			IF Munsch.bSetAirTemp
			THEN
				nWatchdog := 0;
				bDone:= FALSE;                               		(* Program done *)
				bBusy := TRUE;                                  	(* Program busy *)
	
				Munsch.bLockedInterface := TRUE;
				Munsch.bSendExe := FALSE;
	
				IF nAirTemp >= nMinAirTemp
				     AND nAirTemp <= nMaxAirTemp
				THEN
					etMunschExtruder := ET_MunschExtruder_eSetCMD;              (* Next step *)
				ELSE
					udnErrorNo := 1;
	
					etMunschExtruder := ET_MunschExtruder_eError;              (* Next step *)
				END_IF

			ELSE
				etMunschExtruder := ET_MunschExtruder_eError;             (* Next step *)
			END_IF

			Munsch.bSetAirTemp := FALSE;

		ELSIF nWatchdog > 1000
		THEN
			Munsch.bSetAirTemp := FALSE;

			etMunschExtruder := ET_MunschExtruder_eError;             (* Next step *)
		END_IF

	ET_MunschExtruder_eSetCMD:
		Munsch.stMunschCmd.etCommand := ET_MUNSCH_CMD_SETAIRTEMP;
		Munsch.stMunschCmd.nAirTemp := nAirTemp;

		etMunschExtruder := ET_MunschExtruder_eExecuteCMD;              (* Next step *)

	ET_MunschExtruder_eExecuteCMD:
		nWatchdog := nWatchdog + 1;

		Munsch.bSendExe := TRUE;

		IF Munsch.bStringReceived
		THEN
			IF Munsch.stMunschRes.etResponse = ET_MUNSCH_RES_SETAIRTEMP
			     AND Munsch.stMunschCmd.nAirTemp = Munsch.stMunschRes.nAirRefTemp
			THEN
				Munsch.bSendExe := FALSE;

				nWatchdog := 0;

				etMunschExtruder := ET_MunschExtruder_eSetREQ;              (* Next step *)

			END_IF

		ELSIF Munsch.bInterfaceError
			    OR nWatchdog > 1000
		THEN
			Munsch.bSendExe := FALSE;

			udnErrorNo := 2;                     (* Error number *)
			etMunschExtruder := ET_MunschExtruder_eError;              (* Next step *)

		END_IF

	ET_MunschExtruder_eSetREQ:
		Munsch.stMunschCmd.etCommand := ET_MUNSCH_CMD_REQAIRREFTEMP;

		etMunschExtruder := ET_MunschExtruder_eExecuteREQ;              (* Next step *)

	ET_MunschExtruder_eExecuteREQ:
		nWatchdog := nWatchdog + 1;

		Munsch.bSendExe := TRUE;

		IF Munsch.bStringReceived
		THEN
			IF Munsch.stMunschRes.etResponse = ET_MUNSCH_RES_REQAIRREFTEMP
			THEN
				Munsch.nAirRefTemp := Munsch.stMunschRes.nAirRefTemp;

				Munsch.bSendExe := FALSE;

				nWatchdog := 0;
				etMunschExtruder := ET_MunschExtruder_eDone;              (* Next step *)
			END_IF

		ELSIF Munsch.bInterfaceError
			    OR nWatchdog > 1000
		THEN
			Munsch.bSendExe := FALSE;

			udnErrorNo := 3;                     (* Error number *)
			etMunschExtruder := ET_MunschExtruder_eError;              (* Next step *)

		END_IF

	ET_MunschExtruder_eError:
		bBusy := FALSE;						(* Command busy *)
		bError := TRUE;						(* Command error  *)

		etMunschExtruder := ET_MunschExtruder_eNoExecute;

	ET_MunschExtruder_eDone:
		bDone := TRUE;						(* Command done *)
		bBusy := FALSE;						(* Command busy *)

		etMunschExtruder := ET_MunschExtruder_eNoExecute;

	ET_MunschExtruder_eNoExecute:
		IF NOT bExecute
		THEN
			(* Reset outputs *)
			bDone := FALSE;						(* Command done *)
			bBusy := FALSE;						(* Command busy *)
			bError := FALSE;						(* Command error  *)

			nWatchdog := 0;
			Munsch.bLockedInterface := FALSE;

			Munsch.stMunschCmd.etCommand := ET_MUNSCH_CMD_NOCMD;
			Munsch.stMunschRes.etResponse := ET_MUNSCH_RES_NOCMD;

			etMunschExtruder := ET_MunschExtruder_eWaitExecute;
		END_IF
END_CASE;

bAirTempAlarm := Munsch.nAirActTemp > Munsch.nAirRefTemp + nAirTempTolerance
				OR Munsch.nAirActTemp > Munsch.nAirRefTemp - nAirTempTolerance;

END_FUNCTION_BLOCK

// ---- POUs/Tc2 Objects/ExternalHardware/Munsch/FB_MunschExtruder_Extruding.TcPOU
FUNCTION_BLOCK FB_MunschExtruder_Extruding
(*

The function block used to control extruding Munsch extruder

Constructor: 		Patryk Panylo
Company:		E. Riexinger GmbH
Date:			13.10.2015
Version:			1.00

Date:			Revision:		Who:				Comment
dd.mm.yyyy		x.xx			Initials			comment

*)
VAR_INPUT
	(* Input variables / Eingang Variablen *)
	bEnable						:BOOL;						(* Enable FB signal *)
	bStart						:BOOL;						(* Start heating *)
	bStop						:BOOL;						(* Start heating *)
	nExtrudingSpeed				:INT;						(* Extruding speed [%] *)
	rExtrudingSpeedOffset			:REAL;						(* Extruding speed [%] *)
	lrExtrudingSpeedMinV			:LREAL;						(* Extruding speed min [V] 16#0000 = 0 [V] *)
	lrExtrudingSpeedMaxV 		:LREAL;						(* Extruding speed max [V] 16#7FFF = 10 [V], 16#3FFF = 5[V] *)
	lrExtrudingSpeedMin			:LREAL;						(* Extruding speed min [%] *)
	lrExtrudingSpeedMax			:LREAL;						(* Extruding speed max [%] *)
END_VAR
VAR_OUTPUT
	(* Output variables / Ausgang Variablen *)
	bDone						:BOOL;						(* Program done *)
	bBusy						:BOOL;						(* Program busy *)
	bError						:BOOL;						(* Error *)
	udnErrorNo					:UDINT;
END_VAR
VAR_IN_OUT
	(* Input Output variables / Ausgang Variablen *)
	Munsch						:ST_MUNSCH_REF;
END_VAR
VAR
	(* Enummerations *)
	etMunschExtruder				:ET_MunschExtruder;

	(* Variables *)
	nWatchdog					:INT;

	nExtrudingSpeedLimitMax		:INT := 16383;					(* The extruding speed limit (absolute value). Value range in V: 0 ...10, 16#3FFF = 5[V]*)

	(* References *)

	(* Interfaces *)

	(* Instances *)
	fbExtrudingSpeed				:FB_ScalingOffset;
	rtStart						:R_TRIG;
	rtStop						:R_TRIG;

	rtStartEx						:R_TRIG;
	rtStopEx						:R_TRIG;
	bStartEx						:BOOL;
	bStopEx						:BOOL;
END_VAR

IF NOT bEnable
THEN
	bDone := FALSE;					(* Program done *)
	bBusy := FALSE;                                  	(* Program not busy *)
	bError := FALSE;                                 	(* Program not error *)
	udnErrorNo := 0;                                 		(* Error number *)

	Munsch.bExtruding := FALSE;

	RETURN;
END_IF;

(* Scale extruding speed *)
fbExtrudingSpeed(
	bEnable := TRUE,
	lrInput := INT_TO_LREAL(nExtrudingSpeed),
	lrXLowLimit := lrExtrudingSpeedMin,
	lrXUpperLimit := lrExtrudingSpeedMax,
	lrYLowLimit := lrExtrudingSpeedMinV,
	lrYUpperLimit := MIN(lrExtrudingSpeedMaxV, nExtrudingSpeedLimitMax),
	usiPrecision := 2,
	lrOffset := rExtrudingSpeedOffset
);

IF NOT Munsch.bHeat
     OR NOT Munsch.bHeated
     OR NOT Munsch.bExtruding
THEN
	Munsch.nExtrudingSpeed := 0;
	(*bStartEx := FALSE;
	bStopEx := FALSE;*)
ELSE
	(*Munsch.nExtrudingSpeed := LREAL_TO_INT(fbExtrudingSpeed.lrOutputPV);*);
END_IF

(* Wait for triger *)
rtStart(
	CLK := bStart
);

rtStop(
	CLK := bStop
);

(* Wait for triger *)
rtStartEx(
	CLK := Munsch.stMunschCmd.etCommand = ET_MUNSCH_CMD_STARTEXTRUDER
		    AND Munsch.stMunschRes.etResponse = ET_MUNSCH_RES_STARTEXTRUDER
		    AND bBusy
);

rtStopEx(
	CLK := Munsch.stMunschCmd.etCommand = ET_MUNSCH_CMD_STOPEXTRUDER
	  	    AND Munsch.stMunschRes.etResponse = ET_MUNSCH_RES_STOPEXTRUDER
		    AND bBusy
);

IF rtStopEx.Q
THEN
	bStartEx := FALSE;
	bStopEx := TRUE;

ELSIF rtStartEx.Q
THEN
	bStartEx := TRUE;
	bStopEx := FALSE;

END_IF

IF bStopEx
THEN
	Munsch.nExtrudingSpeed := 0;
ELSIF bStartEx
THEN
	Munsch.nExtrudingSpeed := LREAL_TO_INT(fbExtrudingSpeed.lrOutputPV);
END_IF

IF rtStop.Q
THEN
	Munsch.bSetAirTemp := FALSE;
	Munsch.bSetMaterialTemp := FALSE;
	Munsch.bStartHeat := FALSE;
	Munsch.bStopHeat  := FALSE;
	Munsch.bStartExtruding := FALSE;
	Munsch.bStopExtruding  := TRUE;
	Munsch.bReadStatus := FALSE;

	Munsch.nExtrudingSpeed := 0;
END_IF

(* Send command *)
CASE etMunschExtruder OF

	ET_MunschExtruder_eWaitExecute:
		IF rtStop.Q
		    OR Munsch.bStopExtruding
		    OR (nExtrudingSpeed = 0
			   AND Munsch.bExtruding)
		THEN
			nWatchdog := 0;

			Munsch.bSetAirTemp := FALSE;
			Munsch.bSetMaterialTemp := FALSE;
			Munsch.bStartHeat := FALSE;
			Munsch.bStopHeat  := FALSE;
			Munsch.bStartExtruding := FALSE;
			Munsch.bStopExtruding  := TRUE;
			Munsch.bReadStatus := FALSE;

			Munsch.nExtrudingSpeed := 0;

			etMunschExtruder := ET_MunschExtruder_eChkInterface;              (* Next step *)

		ELSIF rtStart.Q
		    	    AND Munsch.bHeat
		             AND Munsch.bHeated
		THEN
			nWatchdog := 0;

			Munsch.bSetAirTemp := FALSE;
			Munsch.bSetMaterialTemp := FALSE;
			Munsch.bStartHeat := FALSE;
			Munsch.bStopHeat  := FALSE;
			Munsch.bStartExtruding := TRUE;
			Munsch.bStopExtruding  := FALSE;
			Munsch.bReadStatus := FALSE;

			etMunschExtruder := ET_MunschExtruder_eChkInterface;              (* Next step *)

		END_IF

	ET_MunschExtruder_eChkInterface:
		nWatchdog := nWatchdog + 1;

		IF NOT Munsch.bLockedInterface
		THEN
			bBusy := FALSE;                                     	(* Program not busy *)
			bError := FALSE;                         		(* Program not error *)
			udnErrorNo := 0;                         		(* Error number *)

			IF Munsch.bStopExtruding
			THEN
				nWatchdog := 0;
				bDone:= FALSE;                               		(* Program done *)
				bBusy := TRUE;                                  	(* Program busy *)
	
				Munsch.nExtrudingSpeed := 0;
	
				Munsch.bLockedInterface := TRUE;
				Munsch.bSendExe := FALSE;
				Munsch.stMunschCmd.etCommand := ET_MUNSCH_CMD_STOPEXTRUDER;
	
				etMunschExtruder := ET_MunschExtruder_eSetCMD;              (* Next step *)
	
			ELSIF Munsch.bStartExtruding
			THEN
				nWatchdog := 0;
				bDone:= FALSE;                               		(* Program done *)
				bBusy := TRUE;                                  	(* Program busy *)
	
				Munsch.nExtrudingSpeed := LREAL_TO_INT(fbExtrudingSpeed.lrOutputPV);
	
				Munsch.bLockedInterface := TRUE;
				Munsch.bSendExe := FALSE;
				Munsch.stMunschCmd.etCommand := ET_MUNSCH_CMD_STARTEXTRUDER;
	
				etMunschExtruder := ET_MunschExtruder_eSetCMD;              (* Next step *)

			ELSE
				etMunschExtruder := ET_MunschExtruder_eError;             (* Next step *)
			END_IF

			Munsch.bStartExtruding := FALSE;
			Munsch.bStopExtruding  := FALSE;

		ELSIF nWatchdog > 1000
		THEN
			Munsch.bStartExtruding := FALSE;
			Munsch.bStopExtruding  := FALSE;

			etMunschExtruder := ET_MunschExtruder_eError;             (* Next step *)
		END_IF

	ET_MunschExtruder_eSetCMD:
		etMunschExtruder := ET_MunschExtruder_eExecuteCMD;              (* Next step *)

	ET_MunschExtruder_eExecuteCMD:
		nWatchdog := nWatchdog + 1;

		Munsch.bSendExe := TRUE;

		IF Munsch.bStringReceived
		THEN
			IF (Munsch.stMunschCmd.etCommand = ET_MUNSCH_CMD_STARTEXTRUDER
			      AND Munsch.stMunschRes.etResponse = ET_MUNSCH_RES_STARTEXTRUDER)
			     OR
			     (Munsch.stMunschCmd.etCommand = ET_MUNSCH_CMD_STOPEXTRUDER
			      AND Munsch.stMunschRes.etResponse = ET_MUNSCH_RES_STOPEXTRUDER)
			THEN
				Munsch.bSendExe := FALSE;

				nWatchdog := 0;
				etMunschExtruder := ET_MunschExtruder_eSetREQ;              (* Next step *)

			END_IF

		ELSIF Munsch.bInterfaceError
			    OR nWatchdog > 1000
		THEN
			Munsch.bSendExe := FALSE;

			udnErrorNo := 1;                     (* Error number *)

			etMunschExtruder := ET_MunschExtruder_eError;              (* Next step *)
		END_IF

	ET_MunschExtruder_eSetREQ:
		Munsch.stMunschCmd.etCommand := ET_MUNSCH_CMD_REQEXTRUDERSTATUS;

		etMunschExtruder := ET_MunschExtruder_eExecuteREQ;              (* Next step *)

	ET_MunschExtruder_eExecuteREQ:
		nWatchdog := nWatchdog + 1;

		Munsch.bSendExe := TRUE;

		IF Munsch.bStringReceived
		THEN
			IF Munsch.stMunschRes.etResponse = ET_MUNSCH_RES_ACKEXTRUDERSTATUSON
			THEN
				Munsch.bExtruding := TRUE;
				Munsch.bSendExe := FALSE;

				nWatchdog := 0;
				etMunschExtruder := ET_MunschExtruder_eDone;              (* Next step *)
			
			ELSIF Munsch.stMunschRes.etResponse = ET_MUNSCH_RES_ACKEXTRUDERSTATUSOFF
			THEN
				Munsch.bExtruding := FALSE;
				Munsch.bSendExe := FALSE;

				nWatchdog := 0;
				etMunschExtruder := ET_MunschExtruder_eDone;              (* Next step *)

			END_IF

		ELSIF Munsch.bInterfaceError
			    OR nWatchdog > 1000
		THEN
			Munsch.bSendExe := FALSE;

			udnErrorNo := 2;                     (* Error number *)

			etMunschExtruder := ET_MunschExtruder_eError;              (* Next step *)
		END_IF

	ET_MunschExtruder_eError:
		bBusy := FALSE;						(* Command busy *)
		bError := TRUE;						(* Command error  *)

		etMunschExtruder := ET_MunschExtruder_eNoExecute;

	ET_MunschExtruder_eDone:
		bDone := TRUE;						(* Command done *)
		bBusy := FALSE;						(* Command busy *)

		etMunschExtruder := ET_MunschExtruder_eNoExecute;

	ET_MunschExtruder_eNoExecute:
		IF NOT bStart
		     AND NOT bStop
		THEN
			(* Reset outputs *)
			bDone := FALSE;						(* Command done *)
			bBusy := FALSE;						(* Command busy *)
			bError := FALSE;						(* Command error  *)

			nWatchdog := 0;
			Munsch.bLockedInterface := FALSE;

			Munsch.stMunschCmd.etCommand := ET_MUNSCH_CMD_NOCMD;
			Munsch.stMunschRes.etResponse := ET_MUNSCH_RES_NOCMD;

			etMunschExtruder := ET_MunschExtruder_eWaitExecute;
		END_IF
END_CASE;

END_FUNCTION_BLOCK

// ---- POUs/Tc2 Objects/ExternalHardware/Munsch/FB_MunschExtruder_Heat.TcPOU
FUNCTION_BLOCK FB_MunschExtruder_Heat
(*

The function block used to control heating Munsch extruder

Constructor: 		Patryk Panylo
Company:		E. Riexinger GmbH
Date:			13.10.2015
Version:			1.00

Date:			Revision:		Who:				Comment
dd.mm.yyyy		x.xx			Initials			comment

*)
VAR_INPUT
	(* Input variables / Eingang Variablen *)
	bEnable						:BOOL;						(* Enable FB signal *)
	bExtruderAirOk				:BOOL;						(* Signal extruder air ok *)
	bStart						:BOOL;						(* Start heating *)
	bStop						:BOOL;						(* Start heating *)
	nMaterialTemp				:INT;						(* Material temperatur *)
	nMinMaterialTemp			:INT;						(* Minimal material temperatur *)
	nMaxMaterialTemp			:INT;						(* Maximal material temperatur *)
	nAirTemp					:INT;						(* Air temperatur *)
	nMinAirTemp					:INT;						(* Minimal air temperatur *)
	nMaxAirTemp				:INT;						(* Maximal air temperatur *)
	tTimeOutAir					:TIME := t#30s;				(* Timeout of air ok *)
END_VAR
VAR_OUTPUT
	(* Output variables / Ausgang Variablen *)
	bExtruderAirOn				:BOOL;						(* Extruder air on*)
	bDone						:BOOL;						(* Program done *)
	bBusy						:BOOL;						(* Program busy *)
	bError						:BOOL;						(* Error *)
	udnErrorNo					:UDINT;
END_VAR
VAR_IN_OUT
	(* Input Output variables / Ausgang Variablen *)
	Munsch						:ST_MUNSCH_REF;
END_VAR
VAR
	(* Enummerations *)
	etMunschExtruder				:ET_MunschExtruder;

	(* Variables *)
	nWatchdog					:INT;

	(* References *)

	(* Interfaces *)

	(* Instances *)
	fbMaterialTemp				:FB_MunschExtruder_MaterialTemp;
	fbAirTemp					:FB_MunschExtruder_AirTemp;
	rtStart						:R_TRIG;
	rtStop						:R_TRIG;
	tonWatchdog					:TON;
END_VAR

IF NOT bEnable
THEN
	bDone := FALSE;					(* Program done *)
	bBusy := FALSE;                                  	(* Program not busy *)
	bError := FALSE;                                 	(* Program not error *)
	udnErrorNo := 0;                                 		(* Error number *)

	fbMaterialTemp(
		bEnable := FALSE,
		Munsch := Munsch
	);

	fbAirTemp(
		bEnable := FALSE,
		Munsch := Munsch
	);

	tonWatchdog(IN := FALSE);

	bExtruderAirOn := FALSE;
	Munsch.bHeat := FALSE;

	RETURN;
END_IF;

(* Wait for triger *)
rtStart(
	CLK := bStart
);

rtStop(
	CLK := bStop
);

IF  NOT Munsch.bHeat
THEN
	Munsch.nExtrudingSpeed := 0;
END_IF

IF rtStop.Q
THEN
	Munsch.bSetAirTemp := FALSE;
	Munsch.bSetMaterialTemp := FALSE;
	Munsch.bStartHeat := FALSE;
	Munsch.bStopHeat  := TRUE;
	Munsch.bStartExtruding := FALSE;
	Munsch.bStopExtruding  := FALSE;
	Munsch.bReadStatus := FALSE;

	Munsch.nExtrudingSpeed := 0;
END_IF

(* Send command *)
CASE etMunschExtruder OF

	ET_MunschExtruder_eWaitExecute:
		IF rtStop.Q
		    OR Munsch.bStopHeat
		THEN
			nWatchdog := 0;

			Munsch.bSetAirTemp := FALSE;
			Munsch.bSetMaterialTemp := FALSE;
			Munsch.bStartHeat := FALSE;
			Munsch.bStopHeat  := TRUE;
			Munsch.bStartExtruding := FALSE;
			Munsch.bStopExtruding  := FALSE;
			Munsch.bReadStatus := FALSE;

			Munsch.nExtrudingSpeed := 0;

			etMunschExtruder := ET_MunschExtruder_eChkInterface;              (* Next step *)

		ELSIF rtStart.Q
		THEN
			nWatchdog := 0;

			Munsch.bSetAirTemp := FALSE;
			Munsch.bSetMaterialTemp := FALSE;
			Munsch.bStartHeat := TRUE;
			Munsch.bStopHeat  := FALSE;
			Munsch.bStartExtruding := FALSE;
			Munsch.bStopExtruding  := FALSE;
			Munsch.bReadStatus := FALSE;

			etMunschExtruder := ET_MunschExtruder_eChkInterface;              (* Next step *)

		END_IF

	ET_MunschExtruder_eChkInterface:
		nWatchdog := nWatchdog + 1;

		IF NOT Munsch.bLockedInterface
		THEN
			bBusy := FALSE;                                     	(* Program not busy *)
			bError := FALSE;                         		(* Program not error *)
			udnErrorNo := 0;                         		(* Error number *)

			IF Munsch.bStopHeat
			THEN
				nWatchdog := 0;
				bDone:= FALSE;                               		(* Program done *)
				bBusy := TRUE;                                  	(* Program busy *)
	
				bExtruderAirOn := FALSE;
				tonWatchdog(IN := FALSE);
	
				Munsch.bLockedInterface := TRUE;
				Munsch.bSendExe := FALSE;
	
				etMunschExtruder := ET_MunschExtruder_eSetCMD;              (* Next step *)
	
			ELSIF Munsch.bStartHeat
			THEN
				nWatchdog := 0;
				bDone:= FALSE;                               		(* Program done *)
				bBusy := TRUE;                                  	(* Program busy *)
	
				fbMaterialTemp(
					bEnable := TRUE,
					bExecute := FALSE,
					nMaterialTemp := nMaterialTemp,
					nMinMaterialTemp := nMinMaterialTemp,
					nMaxMaterialTemp := nMaxMaterialTemp,
					Munsch := Munsch
				);
				
				fbAirTemp(
					bEnable := TRUE,
					bExecute := FALSE,
					nAirTemp := nAirTemp,
					nMinAirTemp := nMinAirTemp,
					nMaxAirTemp := nMaxAirTemp,
					Munsch := Munsch
				);
	
				bExtruderAirOn := TRUE;
				tonWatchdog(IN := FALSE);

				Munsch.bLockedInterface := TRUE;
				Munsch.bSendExe := FALSE;

				etMunschExtruder := ET_MunschExtruder_eSetCMD;              (* Next step *)

			ELSE
				etMunschExtruder :=  ET_MunschExtruder_eError;             (* Next step *)
			END_IF

			Munsch.bStartHeat := FALSE;
			Munsch.bStopHeat  := FALSE;

		ELSIF nWatchdog > 1000
		THEN
			Munsch.bStartHeat := FALSE;
			Munsch.bStopHeat  := FALSE;

			etMunschExtruder :=  ET_MunschExtruder_eError;             (* Next step *)
		END_IF

	ET_MunschExtruder_eSetCMD:
		tonWatchdog(
			IN := TRUE,
			PT:= tTimeOutAir
		);

		IF tonWatchdog.Q
		THEN
			tonWatchdog(IN := FALSE);

			bExtruderAirOn := FALSE;

			udnErrorNo := 1;

			etMunschExtruder := ET_MunschExtruder_eError;             (* Next step *)

		ELSIF bExtruderAirOn
		THEN
			IF bExtruderAirOk
			THEN
				tonWatchdog(IN := FALSE);

				etMunschExtruder := ET_MunschExtruder_eSetMaterialTemp;              (* Next step *)
			END_IF
		ELSE
			Munsch.stMunschCmd.etCommand := ET_MUNSCH_CMD_STOPHEAT;

			tonWatchdog(IN := FALSE);

			etMunschExtruder := ET_MunschExtruder_eExecuteCMD;              (* Next step *)
		END_IF

	ET_MunschExtruder_eSetMaterialTemp:
		nWatchdog := nWatchdog + 1;

		Munsch.bLockedInterface := FALSE;

		fbMaterialTemp(
			bEnable := TRUE,
			bExecute := TRUE,
			nMaterialTemp := nMaterialTemp,
			nMinMaterialTemp := nMinMaterialTemp,
			nMaxMaterialTemp := nMaxMaterialTemp,
			Munsch := Munsch
		);

		IF (NOT fbMaterialTemp.bBusy
		     AND fbMaterialTemp.bError)
		     OR nWatchdog > 1000
		THEN
			fbMaterialTemp(
				bEnable := TRUE,
				bExecute := FALSE,
				Munsch := Munsch
			);

			udnErrorNo := 2;                     (* Error number *)

			etMunschExtruder := ET_MunschExtruder_eError;             (* Next step *)
		
		ELSIF NOT fbMaterialTemp.bBusy
			   AND  fbMaterialTemp.bDone
		THEN
			fbMaterialTemp(
				bEnable := TRUE,
				bExecute := FALSE,
				Munsch := Munsch
			);

			nWatchdog := 0;

			etMunschExtruder := ET_MunschExtruder_eSetAirTemp;             (* Next step *)

		END_IF;

		Munsch.bLockedInterface := TRUE;
		Munsch.bReadStatus := FALSE;

	ET_MunschExtruder_eSetAirTemp:
		nWatchdog := nWatchdog + 1;

		Munsch.bLockedInterface := FALSE;

		fbAirTemp(
			bEnable := TRUE,
			bExecute := TRUE,
			nAirTemp := nAirTemp,
			nMinAirTemp := nMinAirTemp,
			nMaxAirTemp := nMaxAirTemp,
			Munsch := Munsch
		);

		IF (NOT fbAirTemp.bBusy
		     AND fbAirTemp.bError)
		     OR nWatchdog > 1000
		THEN
			fbAirTemp(
				bEnable := TRUE,
				bExecute := FALSE,
				Munsch := Munsch
			);

			udnErrorNo := 3;                     (* Error number *)

			etMunschExtruder := ET_MunschExtruder_eError;             (* Next step *)

		ELSIF NOT fbAirTemp.bBusy
			   AND fbAirTemp.bDone
		THEN
			fbAirTemp(
				bEnable := TRUE,
				bExecute := FALSE,
				Munsch := Munsch
			);

			nWatchdog := 0;

			Munsch.stMunschCmd.etCommand := ET_MUNSCH_CMD_STARTHEAT;

			etMunschExtruder := ET_MunschExtruder_eExecuteCMD;             (* Next step *)
		
		END_IF;

		Munsch.bLockedInterface := TRUE;
		Munsch.bReadStatus := FALSE;

	ET_MunschExtruder_eExecuteCMD:
		nWatchdog := nWatchdog + 1;

		Munsch.bSendExe := TRUE;

		IF Munsch.bStringReceived
		THEN
			IF (bExtruderAirOn
			      AND Munsch.stMunschRes.etResponse = ET_MUNSCH_RES_STARTHEAT)
			     OR
			     (NOT bExtruderAirOn
			      AND Munsch.stMunschRes.etResponse = ET_MUNSCH_RES_STOPHEAT)
			THEN
				Munsch.bSendExe := FALSE;

				nWatchdog := 0;

				etMunschExtruder := ET_MunschExtruder_eSetREQ;              (* Next step *)

			END_IF

		ELSIF Munsch.bInterfaceError
			    OR nWatchdog > 1000
		THEN
			Munsch.bSendExe := FALSE;

			udnErrorNo := 4;                     (* Error number *)

			etMunschExtruder := ET_MunschExtruder_eError;              (* Next step *)

		END_IF

	ET_MunschExtruder_eSetREQ:
		Munsch.stMunschCmd.etCommand := ET_MUNSCH_CMD_REQHEATSTATUS;

		etMunschExtruder := ET_MunschExtruder_eExecuteREQ;              (* Next step *)

	ET_MunschExtruder_eExecuteREQ:
		nWatchdog := nWatchdog + 1;

		Munsch.bSendExe := TRUE;

		IF Munsch.bStringReceived
		THEN
			IF Munsch.stMunschRes.etResponse = ET_MUNSCH_RES_ACKHEATSTATUSON
			THEN
				Munsch.bHeat := TRUE;
				Munsch.bSendExe := FALSE;

				nWatchdog := 0;
				etMunschExtruder := ET_MunschExtruder_eDone;              (* Next step *)
			
			ELSIF Munsch.stMunschRes.etResponse = ET_MUNSCH_RES_ACKHEATSTATUSOFF
			THEN
				Munsch.bHeat := FALSE;
				Munsch.bSendExe := FALSE;

				nWatchdog := 0;
				etMunschExtruder := ET_MunschExtruder_eDone;              (* Next step *)

			END_IF

		ELSIF Munsch.bInterfaceError
			    OR nWatchdog > 1000
		THEN
			Munsch.bSendExe := FALSE;

			udnErrorNo := 5;                     (* Error number *)

			etMunschExtruder := ET_MunschExtruder_eError;              (* Next step *)

		END_IF

	ET_MunschExtruder_eError:
		bBusy := FALSE;						(* Command busy *)
		bError := TRUE;						(* Command error  *)

		etMunschExtruder := ET_MunschExtruder_eNoExecute;

	ET_MunschExtruder_eDone:
		bDone := TRUE;						(* Command done *)
		bBusy := FALSE;						(* Command busy *)

		etMunschExtruder := ET_MunschExtruder_eNoExecute;

	ET_MunschExtruder_eNoExecute:
		IF NOT bStart
		     AND NOT bStop
		THEN
			(* Reset outputs *)
			bDone := FALSE;						(* Command done *)
			bBusy := FALSE;						(* Command busy *)
			bError := FALSE;						(* Command error  *)

			nWatchdog := 0;
			Munsch.bLockedInterface := FALSE;

			Munsch.stMunschCmd.etCommand := ET_MUNSCH_CMD_NOCMD;
			Munsch.stMunschRes.etResponse := ET_MUNSCH_RES_NOCMD;

			etMunschExtruder := ET_MunschExtruder_eWaitExecute;
		END_IF
END_CASE;

END_FUNCTION_BLOCK

// ---- POUs/Tc2 Objects/ExternalHardware/Munsch/FB_MunschExtruder_MaterialTemp.TcPOU
FUNCTION_BLOCK FB_MunschExtruder_MaterialTemp
(*

The function block used to control set material temperature on munschs extruder

Constructor: 		Patryk Panylo
Company:		E. Riexinger GmbH
Date:			18.10.2015
Version:			1.00

Date:			Revision:		Who:				Comment
dd.mm.yyyy		x.xx			Initials			comment

*)
VAR_INPUT
	(* Input variables / Eingang Variablen *)
	bEnable						:BOOL;						(* Enable FB signal *)
	bExecute					:BOOL;						(* Execut the function block *)
	nMaterialTemp				:INT;						(* Material temperatur *)
	nMinMaterialTemp			:INT;						(* Minimal material temperatur *)
	nMaxMaterialTemp			:INT;						(* Maximal material temperatur *)
	nMaterialTempTolerance		:INT := 5;						(* Material temperatur tolerance*)
END_VAR
VAR_OUTPUT
	(* Output variables / Ausgang Variablen *)
	bMaterialTempAlarm			:BOOL;						(* Exceeded material temperature tolerance  *)
	bDone						:BOOL;						(* Program done *)
	bBusy						:BOOL;						(* Program busy *)
	bError						:BOOL;						(* Error *)
	udnErrorNo					:UDINT;
END_VAR
VAR_IN_OUT
	(* Input Output variables / Ausgang Variablen *)
	Munsch						:ST_MUNSCH_REF;
END_VAR
VAR
	(* Enummerations *)
	etMunschExtruder				:ET_MunschExtruder;

	(* Variables *)
	nWatchdog					:INT;

	(* References *)

	(* Interfaces *)

	(* Instances *)
	rtExecute						:R_TRIG;

END_VAR

IF NOT bEnable
THEN
	bDone := FALSE;					(* Program done *)
	bBusy := FALSE;                                  	(* Program not busy *)
	bError := FALSE;                                 	(* Program not error *)
	udnErrorNo := 0;                                 		(* Error number *)

	RETURN;
END_IF;

(* Wait for triger *)
rtExecute(CLK := bExecute);

(* Send command *)
CASE etMunschExtruder OF

	ET_MunschExtruder_eWaitExecute:
		IF rtExecute.Q
		THEN
			nWatchdog := 0;

			Munsch.bSetAirTemp := FALSE;
			Munsch.bSetMaterialTemp := TRUE;
			Munsch.bStartHeat := FALSE;
			Munsch.bStopHeat  := FALSE;
			Munsch.bStartExtruding := FALSE;
			Munsch.bStopExtruding  := FALSE;
			Munsch.bReadStatus := FALSE;

			etMunschExtruder := ET_MunschExtruder_eChkInterface;              (* Next step *)
		END_IF

	ET_MunschExtruder_eChkInterface:
		nWatchdog := nWatchdog + 1;

		IF NOT Munsch.bLockedInterface
		THEN
			bBusy := FALSE;                                     	(* Program not busy *)
			bError := FALSE;                         		(* Program not error *)
			udnErrorNo := 0;                         		(* Error number *)

			IF Munsch.bSetMaterialTemp
			THEN
				nWatchdog := 0;
				bDone:= FALSE;                               		(* Program done *)
				bBusy := TRUE;                                  	(* Program busy *)
	
				Munsch.bLockedInterface := TRUE;
				Munsch.bSendExe := FALSE;
	
				IF nMaterialTemp >= nMinMaterialTemp
				     AND nMaterialTemp <= nMaxMaterialTemp
				THEN
					etMunschExtruder := ET_MunschExtruder_eSetCMD;              (* Next step *)
				ELSE
					udnErrorNo := 1;
	
					etMunschExtruder := ET_MunschExtruder_eError;              (* Next step *)
				END_IF

			ELSE
				etMunschExtruder := ET_MunschExtruder_eError;             (* Next step *)
			END_IF

			Munsch.bSetMaterialTemp := FALSE;

		ELSIF nWatchdog > 1000
		THEN
			Munsch.bSetMaterialTemp := FALSE;

			etMunschExtruder := ET_MunschExtruder_eError;             (* Next step *)
		END_IF

	ET_MunschExtruder_eSetCMD:
		Munsch.stMunschCmd.etCommand := ET_MUNSCH_CMD_SETMATERIALTEMP;
		Munsch.stMunschCmd.nMaterialTemp := nMaterialTemp;

		etMunschExtruder := ET_MunschExtruder_eExecuteCMD;              (* Next step *)

	ET_MunschExtruder_eExecuteCMD:
		nWatchdog := nWatchdog + 1;

		Munsch.bSendExe := TRUE;

		IF Munsch.bStringReceived
		THEN
			IF Munsch.stMunschRes.etResponse = ET_MUNSCH_RES_SETMATERIALTEMP
			     AND Munsch.stMunschCmd.nMaterialTemp = Munsch.stMunschRes.nMaterialRefTemp
			THEN
				Munsch.bSendExe := FALSE;

				nWatchdog := 0;
				etMunschExtruder := ET_MunschExtruder_eSetREQ;              (* Next step *)
			END_IF

		ELSIF Munsch.bInterfaceError
			    OR nWatchdog > 1000
		THEN
			Munsch.bSendExe := FALSE;

			udnErrorNo := 2;                     (* Error number *)
			etMunschExtruder := ET_MunschExtruder_eError;              (* Next step *)
		END_IF

	ET_MunschExtruder_eSetREQ:
		Munsch.stMunschCmd.etCommand := ET_MUNSCH_CMD_REQMATERIALREFTEMP;

		etMunschExtruder := ET_MunschExtruder_eExecuteREQ;              (* Next step *)

	ET_MunschExtruder_eExecuteREQ:
		nWatchdog := nWatchdog + 1;

		Munsch.bSendExe := TRUE;

		IF Munsch.bStringReceived
		THEN
			IF Munsch.stMunschRes.etResponse = ET_MUNSCH_RES_REQMATERIALREFTEMP
			THEN
				Munsch.nMaterialRefTemp := Munsch.stMunschRes.nMaterialRefTemp;

				Munsch.bSendExe := FALSE;

				nWatchdog := 0;
				etMunschExtruder := ET_MunschExtruder_eDone;              (* Next step *)

			END_IF

		ELSIF Munsch.bInterfaceError
			    OR nWatchdog > 1000
		THEN
			Munsch.bSendExe := FALSE;

			udnErrorNo := 3;                     (* Error number *)
			etMunschExtruder := ET_MunschExtruder_eError;              (* Next step *)
		END_IF

	ET_MunschExtruder_eError:
		bBusy := FALSE;						(* Command busy *)
		bError := TRUE;						(* Command error  *)

		etMunschExtruder := ET_MunschExtruder_eNoExecute;

	ET_MunschExtruder_eDone:
		bDone := TRUE;						(* Command done *)
		bBusy := FALSE;						(* Command busy *)

		etMunschExtruder := ET_MunschExtruder_eNoExecute;

	ET_MunschExtruder_eNoExecute:
		IF NOT bExecute
		THEN
			(* Reset outputs *)
			bDone := FALSE;						(* Command done *)
			bBusy := FALSE;						(* Command busy *)
			bError := FALSE;						(* Command error  *)

			nWatchdog := 0;
			Munsch.bLockedInterface := FALSE;

			Munsch.stMunschCmd.etCommand := ET_MUNSCH_CMD_NOCMD;
			Munsch.stMunschRes.etResponse := ET_MUNSCH_RES_NOCMD;

			etMunschExtruder := ET_MunschExtruder_eWaitExecute;
		END_IF
END_CASE;

bMaterialTempAlarm := Munsch.nMaterialActTemp > Munsch.nMaterialRefTemp + nMaterialTempTolerance
					 OR Munsch.nMaterialActTemp > Munsch.nMaterialRefTemp - nMaterialTempTolerance;

END_FUNCTION_BLOCK

// ---- POUs/Tc2 Objects/ExternalHardware/Munsch/FB_MunschExtruder_ReadStatus.TcPOU
FUNCTION_BLOCK FB_MunschExtruder_ReadStatus
(*

The function block used to read status of Munsch extruder

Constructor: 		Patryk Panylo
Company:		E. Riexinger GmbH
Date:			13.10.2015
Version:			1.00

Date:			Revision:		Who:				Comment
dd.mm.yyyy		x.xx			Initials			comment

*)
VAR_INPUT
	(* Input variables / Eingang Variablen *)
	bEnable						:BOOL;						(* Enable FB signal *)
	bExecute					:BOOL;						(* Execute read status *)
	tReadStatus					:TIME := t#0ms;				(* Read current status *)
END_VAR
VAR_OUTPUT
	(* Output variables / Ausgang Variablen *)
	bDone						:BOOL;						(* Program done *)
	bBusy						:BOOL;						(* Program busy *)
	bError						:BOOL;						(* Error *)
	udnErrorNo					:UDINT;
END_VAR
VAR_IN_OUT
	(* Input Output variables / Ausgang Variablen *)
	Munsch						:ST_MUNSCH_REF;
END_VAR
VAR
	(* Enummerations *)
	etMunschExtruder				:ET_MunschExtruder;

	(* Variables *)
	bReadStatus					:BOOL;
	nReqCount					:INT;
	nWatchdog					:INT;

	(* References *)

	(* Interfaces *)

	(* Instances *)
	tonReadStatus				:TON;
	rtExecute						:R_TRIG;
	rtStart						:R_TRIG;
	rtStop						:R_TRIG;
END_VAR

IF NOT bEnable
THEN
	bDone := FALSE;					(* Program done *)
	bBusy := FALSE;                                  	(* Program not busy *)
	bError := FALSE;                                 	(* Program not error *)
	udnErrorNo := 0;                                 		(* Error number *)

	tonReadStatus(
		IN := FALSE,
	);

	RETURN;
END_IF;

rtStart(CLK := (tReadStatus > t#0ms
		       OR  (bExecute AND tReadStatus = t#0ms))
		       AND NOT Munsch.bLockedInterface);
rtStop(CLK := tReadStatus = t#0ms);

IF rtStop.Q
THEN
	Munsch.bReadStatus := FALSE;

ELSIF rtStart.Q
THEN
	Munsch.bReadStatus := TRUE;

	bDone := FALSE;					(* Program done *)
	bBusy := FALSE;                                  	(* Program not busy *)
	bError := FALSE;                                 	(* Program not error *)
	udnErrorNo := 0;                                 		(* Error number *)

	etMunschExtruder := ET_MunschExtruder_eWaitExecute;              (* Next step *)

END_IF

tonReadStatus(
	IN := Munsch.bReadStatus,
	PT := tReadStatus,
);

rtExecute(
	CLK := tonReadStatus.Q
);

(* Send command *)
CASE etMunschExtruder OF

	ET_MunschExtruder_eWaitExecute:
		bBusy := FALSE;                                     	(* Program not busy *)
		bError := FALSE;                         		(* Program not error *)
		udnErrorNo := 0;                         		(* Error number *)

		IF rtExecute.Q
		     AND NOT Munsch.bLockedInterface
		THEN
			nWatchdog := 0;
			bDone:= FALSE;                               		(* Program done *)
			bBusy := TRUE;                                  	(* Program busy *)

			nReqCount  := 0;
			Munsch.bLockedInterface := TRUE;
			Munsch.bSendExe := FALSE;

			etMunschExtruder := ET_MunschExtruder_eSetREQ;              (* Next step *)

		END_IF

	ET_MunschExtruder_eSetREQ:
		CASE nReqCount
		OF
			0: Munsch.stMunschCmd.etCommand := ET_MUNSCH_CMD_REQHEATSTATUS;
			    nReqCount := 1;
			1: Munsch.stMunschCmd.etCommand := ET_MUNSCH_CMD_REQEXTRUDERSTATUS;
			    nReqCount := 2;
			2: Munsch.stMunschCmd.etCommand := ET_MUNSCH_CMD_REQMATERIALREFTEMP;
			    nReqCount := 3;
			3: Munsch.stMunschCmd.etCommand := ET_MUNSCH_CMD_REQMATERIALACTTEMP;
			    nReqCount := 4;
			4: Munsch.stMunschCmd.etCommand := ET_MUNSCH_CMD_REQAIRREFTEMP;
			    nReqCount := 5;
			5: Munsch.stMunschCmd.etCommand := ET_MUNSCH_CMD_REQAIRACTTEMP;
			    nReqCount := 6;
			6: Munsch.stMunschCmd.etCommand := ET_MUNSCH_CMD_REQSTATUS;
				nReqCount := 0;
		END_CASE

		etMunschExtruder := ET_MunschExtruder_eExecuteREQ;              (* Next step *)

	ET_MunschExtruder_eExecuteREQ:
		nWatchdog := nWatchdog + 1;

		Munsch.bSendExe := TRUE;

		IF Munsch.bStringReceived
		THEN
			IF Munsch.stMunschRes.etResponse = ET_MUNSCH_RES_ACKHEATSTATUSON
			THEN
				Munsch.bHeat := TRUE;
				Munsch.bSendExe := FALSE;

				nWatchdog := 0;
				IF nReqCount > 0
				     AND Munsch.bReadStatus
				THEN
					etMunschExtruder := ET_MunschExtruder_eSetREQ;
				ELSE
					etMunschExtruder := ET_MunschExtruder_eDone;              (* Next step *)
				END_IF
			
			ELSIF Munsch.stMunschRes.etResponse = ET_MUNSCH_RES_ACKHEATSTATUSOFF
			THEN
				Munsch.bHeat := FALSE;
				Munsch.bSendExe := FALSE;

				nWatchdog := 0;
				IF nReqCount > 0
				    AND Munsch.bReadStatus
				THEN
					etMunschExtruder := ET_MunschExtruder_eSetREQ;
				ELSE
					etMunschExtruder := ET_MunschExtruder_eDone;              (* Next step *)
				END_IF

			ELSIF Munsch.stMunschRes.etResponse = ET_MUNSCH_RES_ACKEXTRUDERSTATUSON
			THEN
				Munsch.bExtruding := TRUE;
				Munsch.bSendExe := FALSE;

				nWatchdog := 0;
				IF nReqCount > 0
				    AND Munsch.bReadStatus
				THEN
					etMunschExtruder := ET_MunschExtruder_eSetREQ;
				ELSE
					etMunschExtruder := ET_MunschExtruder_eDone;              (* Next step *)
				END_IF
			
			ELSIF Munsch.stMunschRes.etResponse = ET_MUNSCH_RES_ACKEXTRUDERSTATUSOFF
			THEN
				Munsch.bExtruding := FALSE;
				Munsch.bSendExe := FALSE;

				nWatchdog := 0;
				IF nReqCount > 0
				     AND Munsch.bReadStatus
				THEN
					etMunschExtruder := ET_MunschExtruder_eSetREQ;
				ELSE
					etMunschExtruder := ET_MunschExtruder_eDone;              (* Next step *)
				END_IF

			ELSIF Munsch.stMunschRes.etResponse = ET_MUNSCH_RES_REQMATERIALREFTEMP
			THEN
				Munsch.nMaterialRefTemp := Munsch.stMunschRes.nMaterialRefTemp;
				Munsch.bSendExe := FALSE;

				nWatchdog := 0;
				IF nReqCount > 0
				     AND Munsch.bReadStatus
				THEN
					etMunschExtruder := ET_MunschExtruder_eSetREQ;
				ELSE
					etMunschExtruder := ET_MunschExtruder_eDone;              (* Next step *)
				END_IF

			ELSIF Munsch.stMunschRes.etResponse = ET_MUNSCH_RES_REQMATERIALACTTEMP
			THEN
				Munsch.nMaterialActTemp := Munsch.stMunschRes.nMaterialActTemp;
				Munsch.bSendExe := FALSE;

				nWatchdog := 0;
				IF nReqCount > 0
				     AND Munsch.bReadStatus
				THEN
					etMunschExtruder := ET_MunschExtruder_eSetREQ;
				ELSE
					etMunschExtruder := ET_MunschExtruder_eDone;              (* Next step *)
				END_IF

			ELSIF Munsch.stMunschRes.etResponse = ET_MUNSCH_RES_REQAIRREFTEMP
			THEN
				Munsch.nAirRefTemp := Munsch.stMunschRes.nAirRefTemp;
				Munsch.bSendExe := FALSE;

				nWatchdog := 0;
				IF nReqCount > 0
				     AND Munsch.bReadStatus
				THEN
					etMunschExtruder := ET_MunschExtruder_eSetREQ;
				ELSE
					etMunschExtruder := ET_MunschExtruder_eDone;              (* Next step *)
				END_IF

			ELSIF Munsch.stMunschRes.etResponse = ET_MUNSCH_RES_REQAIRACTTEMP
			THEN
				Munsch.nAirActTemp := Munsch.stMunschRes.nAirActTemp;
				Munsch.bSendExe := FALSE;

				nWatchdog := 0;
				IF nReqCount > 0
				     AND Munsch.bReadStatus
				THEN
					etMunschExtruder := ET_MunschExtruder_eSetREQ;
				ELSE
					etMunschExtruder := ET_MunschExtruder_eDone;              (* Next step *)
				END_IF

			ELSIF Munsch.stMunschRes.etResponse = ET_MUNSCH_RES_REQSTATUSHEATED
			THEN
				Munsch.bHeating := FALSE;
				Munsch.bHeated := TRUE;
				Munsch.bError := FALSE;
				Munsch.bSendExe := FALSE;

				nWatchdog := 0;
				IF nReqCount > 0
				     AND Munsch.bReadStatus
				THEN
					etMunschExtruder := ET_MunschExtruder_eSetREQ;
				ELSE
					etMunschExtruder := ET_MunschExtruder_eDone;              (* Next step *)
				END_IF

			ELSIF Munsch.stMunschRes.etResponse = ET_MUNSCH_RES_REQSTATUSHEATING
			THEN
				Munsch.bHeating := Munsch.bHeat;
				Munsch.bHeated := FALSE;
				Munsch.bError := FALSE;
				Munsch.bSendExe := FALSE;

				nWatchdog := 0;
				IF nReqCount > 0
				     AND Munsch.bReadStatus
				THEN
					etMunschExtruder := ET_MunschExtruder_eSetREQ;
				ELSE
					etMunschExtruder := ET_MunschExtruder_eDone;              (* Next step *)
				END_IF

			ELSIF Munsch.stMunschRes.etResponse = ET_MUNSCH_RES_REQSTATUSERROR
			THEN
				Munsch.bHeating := FALSE;
				Munsch.bHeated := FALSE;
				Munsch.bError := TRUE;
				Munsch.bSendExe := FALSE;

				nWatchdog := 0;
				IF nReqCount > 0
				     AND Munsch.bReadStatus
				THEN
					etMunschExtruder := ET_MunschExtruder_eSetREQ;
				ELSE
					etMunschExtruder := ET_MunschExtruder_eDone;              (* Next step *)
				END_IF

			END_IF

		ELSIF Munsch.bInterfaceError
 			    OR nWatchdog > 1000
		THEN
			Munsch.bSendExe := FALSE;

			udnErrorNo := 2;                     (* Error number *)

			etMunschExtruder := ET_MunschExtruder_eError;              (* Next step *)
		END_IF

	ET_MunschExtruder_eError:
		bBusy := FALSE;						(* Command busy *)
		bError := TRUE;						(* Command error  *)

		etMunschExtruder := ET_MunschExtruder_eNoExecute;

	ET_MunschExtruder_eDone:
		bDone := TRUE;						(* Command done *)
		bBusy := FALSE;						(* Command busy *)

		etMunschExtruder := ET_MunschExtruder_eNoExecute;

	ET_MunschExtruder_eNoExecute:
		IF tReadStatus > t#0ms
		THEN
			tonReadStatus(
				IN := FALSE,
				PT := tReadStatus,
			);
		END_IF

		IF NOT tonReadStatus.Q
		     OR (NOT bExecute AND tReadStatus = t#0ms)
		THEN
			(* Reset outputs *)
			bDone := FALSE;						(* Command done *)
			bBusy := FALSE;						(* Command busy *)
			bError := FALSE;						(* Command error  *)

			nWatchdog := 0;
			Munsch.bLockedInterface := FALSE;

			IF tReadStatus = t#0ms
			THEN
				Munsch.bReadStatus := FALSE;
			END_IF

			etMunschExtruder := ET_MunschExtruder_eWaitExecute;
		END_IF
END_CASE;

END_FUNCTION_BLOCK

// ---- POUs/Tc2 Objects/ExternalHardware/Munsch/FB_MUNSCH_EXTRUDER_REF.TcPOU
FUNCTION_BLOCK FB_MUNSCH_EXTRUDER_REF
VAR_INPUT
	bSendExe					:BOOL;						(* Send execute *)
	tSendPeriod					:TIME := t#0s;					(* Send data every period. If tSendPeriod is 0 then th function is not active *)
	bLockedInterface				:BOOL;						(* Locked interface *)
	bHeat						:BOOL;						(* Heat status ON = TRUE, OFF = FALSE *)
	bHeating						:BOOL;						(* Heating status ON = TRUE, OFF = FALSE *)
	bHeated						:BOOL;						(* Heated status ON = TRUE, OFF = FALSE *)
	bError						:BOOL;						(* Error ON = TRUE, OFF = FALSE *)
	bExtruding					:BOOL;						(* Extruder status ON = TRUE, OFF = FALSE *)
	nMaterialRefTemp			:INT;						(* Referenc material temperature *)
	nMaterialActTemp				:INT;						(* Current material temperature *)
	nAirRefTemp					:INT;						(* Referenc air temperature *)
	nAirActTemp					:INT;						(* Current air temperature *)
	stMunschCmd				:ST_MUNSCH_CMD_Data;
	stMunschRes					:ST_MUNSCH_RES_Data;
	bInterfaceReady				:BOOL;						(* Interface ready to use *)
	bInterfaceError				:BOOL;						(* Interface error *)
	bStringReceived				:BOOL;						(* String received *)
	bSetAirTemp					:BOOL;						(* Set air temperature *)
	bSetMaterialTemp			:BOOL;						(* Set material temperature *)
	bStartHeat					:BOOL;						(* Heat start *)
	bStopHeat					:BOOL;						(* Heat stop *)
	bStartExtruding				:BOOL;						(* Extruding start *)
	bStopExtruding				:BOOL;						(* Extruding start *)
	bReadStatus					:BOOL;						(* Enable read current status *)
	bExtrudingStop				:BOOL;						(* Extruding stop *)
	nExtrudingSpeed				:INT;						(* Extruding speed *)
END_VAR
VAR_OUTPUT

END_VAR
VAR_IN_OUT

END_VAR
VAR

END_VAR

;

END_FUNCTION_BLOCK

// ---- POUs/Tc2 Objects/ExternalHardware/YASKAWA/FB_YASKAWA_Controller.TcPOU
FUNCTION_BLOCK FB_YASKAWA_Controller
(*

The function block used to control axis.

Constructor: 		Patryk Panylo
Company:		E. Riexinger GmbH
Date:			20.06.2018
Version:			1.00

Date:			Revision:		Who:				Comment
dd.mm.yyyy		x.xx			Initials			comment

*)
VAR_INPUT
	(* Input variables / Eingang Variablen *)
	bEnable						:BOOL;						(* Signal FB enable *)
	etMachineMode				:ET_MachineMode;			(* Machine mode *)
	etMachineState				:ET_MachineState;			(* Machine state *)
	bDrivesOn					:BOOL;						(* Enable the drives *)
	bMoveOn					:BOOL;						(* Enable the move enable *)
	bReset						:BOOL;						(* Signal reset *)
	bExeReset					:BOOL;						(* Execute auto reset *)
	lrOverride					:LREAL;						(* Override 100% percent *)
END_VAR
VAR_OUTPUT
	(* Output variables / Ausgang Variablen *)
	bStatus						:BOOL;						(* Feedback *)
	bStatusDelay					:BOOL;						(* Feedback delay *)
	bReseted					:BOOL;						(* Reset completed *)
	bError						:BOOL;						(* Controller error *)
	udnErrorNo					:UDINT;						(* Error number *)
	bInHome						:BOOL;						(* In home *)
	bNotMoving					:BOOL;						(* Status of moving *)
	bNotInCrashAreaMachine		:BOOL;						(* Status not in crash area *)
END_VAR
VAR_IN_OUT
	(* Input Output variables / Ausgang Variablen *)
	Yaskawa					:ST_YASKAWA_REF;				(* The YASKAWA_REF data type  is an interface between the PLC and the YASKAWA and contains axis information *)
END_VAR
VAR
	(* Enummerations *)

	(* Variables *)
	tStatusDelay					:TIME := t#1s;					(* Status delay time *)

	bFirstTime					:BOOL;

	(* References *)

	(* Interfaces *)

	(* Instances *)
	fbPower						:FB_YASKAWA_Power;		(* The function block is used to enable for an axis *)
	tonStatusDelay				:TON;						(* Delay controller enabled status *)
	fbReset						:FB_YASKAWA_Reset;			(* An axis reset is carried out with the function block *)

END_VAR


IF NOT bEnable							(* Signal FB enable *)
THEN
	bStatus := FALSE;						(* Feedback *)
	bStatusDelay := FALSE;				(* Feedback *)
	bError := FALSE;						(* Controller error *)
	udnErrorNo := 0;						(* Error number *)

	bFirstTime := FALSE;
	RETURN;
END_IF

IF NOT bFirstTime
THEN

	bFirstTime := TRUE;
END_IF;

A_Power();
A_Reset();
A_Error();

(* In home *)
bInHome := Yaskawa.stYaskawaToPlc.bInHome;

(* Status not moving *)
bNotMoving := Yaskawa.stYaskawaToPlc.bNotMoving;

(* Status not in crash area *)
bNotInCrashAreaMachine := Yaskawa.stYaskawaToPlc.bNotInCrashAreaMachine;

ACTION A_Error:

bError := fbReset.bError
	         OR fbPower.bError;
END_ACTION

ACTION A_Power:

fbPower(
	bEnable := TRUE,
	bAutoHand := etMachineMode = ET_MachineMode_eHome
			         OR etMachineMode = ET_MachineMode_eStepping
			         OR etMachineMode = ET_MachineMode_eAutomatic,
	bDrivesOn :=  bDrivesOn,
	bMoveOn := bMoveOn,
	lrOverride := lrOverride,
	Yaskawa := Yaskawa
 );

tonStatusDelay(
	IN := fbPower.bStatus,
	PT := SEL(etMachineMode = ET_MachineMode_eManual, tStatusDelay, t#0ms),
	Q => bStatusDelay
);
END_ACTION

ACTION A_Reset:

fbReset(
	bExecute := bReset
	            	     XOR bExeReset,
	Yaskawa := Yaskawa,
	bDone => bReseted
);
END_ACTION

END_FUNCTION_BLOCK

// ---- POUs/Tc2 Objects/ExternalHardware/YASKAWA/FB_YASKAWA_Power.TcPOU
FUNCTION_BLOCK FB_YASKAWA_Power
(*

The function block used to enable drives for an yaskawa

Constructor: 		Patryk Panylo
Company:		E. Riexinger GmbH
Date:			20.06.2018
Version:			1.00

Date:			Revision:		Who:				Comment

*)
VAR_INPUT
	(* Input variables / Eingang Variablen *)
	bEnable						:BOOL;			(* Signal FB enable *)
	bAutoHand					:BOOL;			(* Auto := TRUE, Hand := FALSE *)
	bDrivesOn					:BOOL;			(* Enable the drives *)
	bMoveOn					:BOOL;			(* Enable the move enable *)
	lrOverride					:LREAL;			(* Velocity override in % for all motion commands. (0 <= Override <= 100.0) *)
END_VAR
VAR_OUTPUT
	(* Output variables / Ausgang Variablen *)
	bStatus						:BOOL;			(* Status = TRUE indicates that the axis is ready for operation. *)
	bError						:BOOL;			(* Error *)
	udnErrorNo					:UDINT;			(* Error number *)
	sErrorMsg					:STRING; 		(* Error message *)
END_VAR
VAR_IN_OUT
	(* Input Output variables / Ausgang Variablen *)
	Yaskawa					:ST_YASKAWA_REF;				(* The YASKAWA_REF data type  is an interface between the PLC and the YASKAWA and contains axis information *)
END_VAR
VAR
	(* Enummerations *)

	(* Variables *)
	tStatusDelay 					:TIME := t#300ms;

	(* References *)

	(* Interfaces *)

	(* Instances *)
	tonStatusDelay				:TON;
END_VAR


IF NOT bEnable
THEN
	Yaskawa.stPlcToYaskawa.bExternalServoOn := FALSE;                   		 (* Switch on *)
	tonStatusDelay(IN := FALSE,
				    PT := tStatusDelay);
ELSE

	IF NOT bDrivesOn
	     OR Yaskawa.stYaskawaToPlc.bAlarmErrorOccured
	THEN
		Yaskawa.stPlcToYaskawa.bCallMasterJob := FALSE;
		Yaskawa.stPlcToYaskawa.bExternalStart := FALSE;
		Yaskawa.stPlcToYaskawa.bExternalHold := FALSE;
		Yaskawa.stPlcToYaskawa.bExternalServoOn := FALSE;						 (* Switch on *)
		Yaskawa.stPlcToYaskawa.bExternalServoOffEStop := TRUE;                   		 (* Switch off *)
		Yaskawa.stPlcToYaskawa.bExternalServoOffHoldStop := FALSE;                   		 (* Switch off *)
	ELSE
		IF bAutoHand			(* Auto *)
		THEN
			IF bMoveOn
			     AND Yaskawa.stYaskawaToPlc.bRemoteModeSelected
			THEN
				Yaskawa.stPlcToYaskawa.bExternalServoOn := TRUE;                   				 (* Switch on *)
				Yaskawa.stPlcToYaskawa.bExternalServoOffEStop := FALSE;                   		 (* Switch off *)
				Yaskawa.stPlcToYaskawa.bExternalServoOffHoldStop := FALSE;                   		 (* Switch off *)
			ELSE
				Yaskawa.stPlcToYaskawa.bExternalServoOn := FALSE;                   				(* Switch on *)
				Yaskawa.stPlcToYaskawa.bExternalServoOffEStop := FALSE;                   		(* Switch off *)
				Yaskawa.stPlcToYaskawa.bExternalServoOffHoldStop := TRUE;				(* Switch off *)
			END_IF
		ELSE				(* Manual *)
			Yaskawa.stPlcToYaskawa.bCallMasterJob := FALSE;
			Yaskawa.stPlcToYaskawa.bExternalStart := FALSE;
			Yaskawa.stPlcToYaskawa.bExternalHold := FALSE;
			Yaskawa.stPlcToYaskawa.bExternalServoOn := FALSE;						(* Switch on *)
			Yaskawa.stPlcToYaskawa.bExternalServoOffEStop := FALSE;                   		(* Switch off *)
			Yaskawa.stPlcToYaskawa.bExternalServoOffHoldStop := FALSE;				(* Switch off *)
		END_IF
	END_IF;
END_IF;

Yaskawa.stPlcToYaskawa.usnOverride := LREAL_TO_USINT(LIMIT(1,lrOverride,100));

tonStatusDelay(IN := Yaskawa.stYaskawaToPlc.bServoIsOn,		(* Control enabled *)
			   PT := tStatusDelay);
bStatus := tonStatusDelay.Q;

END_FUNCTION_BLOCK

// ---- POUs/Tc2 Objects/ExternalHardware/YASKAWA/FB_YASKAWA_Reset.TcPOU
FUNCTION_BLOCK FB_YASKAWA_Reset
(*

The function block used to reset the yaskawa message.

Constructor: 		Patryk Panylo
Company:		E. Riexinger GmbH
Date:			20.06.2018
Version:			1.00

Date:			Revision:		Who:				Comment

*)
VAR_INPUT
	(* Input variables / Eingang Variablen *)
	bExecute					:BOOL;		(* Execut the function block *)
	bExtReset					:BOOL;
END_VAR
VAR_OUTPUT
	(* Output variables / Ausgang Variablen *)
	bDone						:BOOL;			(* Program done. *)
	bBusy						:BOOL;			(* Program busy *)
	bError						:BOOL;			(* Error *)
	udnErrorNo					:UDINT;			(* Error number *)
	sErrorMsg					:STRING; 		(* Error message *)
END_VAR
VAR_IN_OUT
	(* Input Output variables / Ausgang Variablen *)
	Yaskawa					:ST_YASKAWA_REF;				(* The YASKAWA_REF data type  is an interface between the PLC and the YASKAWA and contains axis information *)
END_VAR
VAR
	(* Enummerations *)

	(* Variables *)

	(* References *)

	(* Interfaces *)

	(* Instances *)
	rtExecute						:R_TRIG;
	rtExtReset					:R_TRIG;
	rtDrivesOn					:R_TRIG;

END_VAR


rtExecute(CLK := bExecute
			      AND Yaskawa.stYaskawaToPlc.bAlarmErrorOccured);
rtDrivesOn(CLK := Yaskawa.stYaskawaToPlc.bServoIsOn
	   		        AND Yaskawa.stPlcToYaskawa.bExternalServoOn);

IF rtExecute.Q
     OR (rtDrivesOn.Q
	    AND Yaskawa.stYaskawaToPlc.bAlarmErrorOccured)
THEN
	bBusy := TRUE;
	Yaskawa.stPlcToYaskawa.bAlarmReset := TRUE;

ELSIF Yaskawa.stPlcToYaskawa.bAlarmReset
	   AND NOT Yaskawa.stYaskawaToPlc.bAlarmErrorOccured
THEN
	bBusy := FALSE;
	Yaskawa.stPlcToYaskawa.bAlarmReset := FALSE;
END_IF;

bDone := bExecute
		AND NOT bBusy
		AND NOT Yaskawa.stYaskawaToPlc.bAlarmErrorOccured;        (* Error *)

END_FUNCTION_BLOCK

// ---- POUs/Tc2 Objects/ExternalHardware/YASKAWA/FB_YASKAWA_REF.TcPOU
FUNCTION_BLOCK FB_YASKAWA_REF
VAR_INPUT
	stYaskawaToPlc				:ST_YASKAWATOPLC;
	stPlcToYaskawa				:ST_PLCTOYASKAWA;

	stTerminalState				AT %I*:ST_TerminalState;
	stRobotToPlc					AT %I*:ST_ROBOTTOPLC;
	stPlcToRobot					AT %Q*:ST_PLCTOROBOT;
END_VAR
VAR_OUTPUT

END_VAR
VAR_IN_OUT

END_VAR
VAR

END_VAR

;

END_FUNCTION_BLOCK

// ---- POUs/Tc2 Objects/ExternalHardware/YASKAWA/FB_YASKAWA_StartPrg.TcPOU
FUNCTION_BLOCK FB_YASKAWA_StartPrg
(*

The function block used to start kuka

Constructor: 		Patryk Panylo
Company:		E. Riexinger GmbH
Date:			18.11.2016
Version:			1.00

Date:			Revision:		Who:				Comment

*)
VAR_INPUT
	(* Input variables / Eingang Variablen *)
	bEnable						:BOOL;			(* Signal FB enable *)
	bReset						:BOOL;			(* Signal reset *)
	bAutoHand					:BOOL;			(* Auto := TRUE, Hand := FALSE *)
	bStart						:BOOL;			(* Start program *)
	bStop						:BOOL;			(* Stop program *)
	bInterrupt						:BOOL;			(* Interrupt *)
	nPrgNo						:INT;			(* Program number *)
END_VAR
VAR_OUTPUT
	(* Output variables / Ausgang Variablen *)
	bRunning					:BOOL;						(* Program running *)
	bDone						:BOOL;						(* Program done *)
	bInterrupted					:BOOL;						(* Program interrupted *)
	bBusy						:BOOL;						(* Program busy *)
	bError						:BOOL;						(* Error *)
	udnErrorNo					:UDINT;
END_VAR
VAR_IN_OUT
	(* Input Output variables / Ausgang Variablen *)
	Yaskawa					:ST_YASKAWA_REF;				(* The YASKAWA_REF data type  is an interface between the PLC and the YASKAWA and contains axis information *)
END_VAR
VAR
	(* Enummerations *)
	etYaskawaStart				:ET_YaskawaStart;

	(* Variables *)
	wDoneFlag					:WORD;
	bFirstTime					:BOOL;

	nWatchdog					:INT;

	(* References *)

	(* Interfaces *)

	(* Instances *)
	rtStart						:R_TRIG;
	rtStop						:R_TRIG;
	rtReset						:R_TRIG;
	rtInterrupt						:R_TRIG;
	tonWatchdog					:TON;

END_VAR


IF NOT bEnable
THEN
	bDone := FALSE;					(* Program done *)
	bInterrupted := FALSE;				(* Program interrupted *)
	bBusy := FALSE;                                  	(* Program not busy *)
	bError := FALSE;                                 	(* Program not error *)
	udnErrorNo := 0;                                 		(* Error number *)

	Yaskawa.stPlcToYaskawa.bCallMasterJob := FALSE;
	Yaskawa.stPlcToYaskawa.bExternalStart := FALSE;
	Yaskawa.stPlcToYaskawa.bExternalHold := FALSE;

	RETURN;
END_IF;

IF NOT bFirstTime
THEN
	tonWatchdog(IN := FALSE);

	Yaskawa.stPlcToYaskawa.bCallMasterJob := FALSE;
	Yaskawa.stPlcToYaskawa.bExternalStart := FALSE;
	Yaskawa.stPlcToYaskawa.bExternalHold := FALSE;

	etYaskawaStart := ET_YaskawaStart_eWaitExecute;              (* Next step *)

	bFirstTime := TRUE;
END_IF

rtReset(CLK := bReset);

IF rtReset.Q
     AND bError
THEN
	bError := FALSE;

	tonWatchdog(IN := FALSE);

	Yaskawa.stPlcToYaskawa.bCallMasterJob := FALSE;
	Yaskawa.stPlcToYaskawa.bExternalStart := FALSE;
	Yaskawa.stPlcToYaskawa.bExternalHold := FALSE;

	etYaskawaStart := ET_YaskawaStart_eWaitExecute;              (* Next step *)
END_IF

rtInterrupt(CLK := bInterrupt);
IF rtInterrupt.Q
THEN
	tonWatchdog(IN := FALSE);

	Yaskawa.stPlcToYaskawa.bCallMasterJob := FALSE;
	Yaskawa.stPlcToYaskawa.bExternalStart := FALSE;
	Yaskawa.stPlcToYaskawa.bExternalHold := FALSE;

	etYaskawaStart := ET_YaskawaStart_eInterrupted;              (* Next step *)
END_IF;

(* Wait for triger *)
rtStart(
	CLK := bStart
);

IF rtStart.Q
     AND NOT bStop
     AND Yaskawa.stYaskawaToPlc.bServoIsOn
     AND NOT Yaskawa.stYaskawaToPlc.bAlarmErrorOccured
THEN
	Yaskawa.stPlcToYaskawa.bCallMasterJob := FALSE;
	Yaskawa.stPlcToYaskawa.bExternalStart := FALSE;

	IF bAutoHand
	THEN
		Yaskawa.stPlcToYaskawa.bExternalHold := FALSE;
	END_IF

	etYaskawaStart := ET_YaskawaStart_eWaitExecute;              (* Next step *)

END_IF

rtStop(
	CLK := bStop
);

IF rtStop.Q
     OR Yaskawa.stYaskawaToPlc.bAlarmErrorOccured
THEN
	Yaskawa.stPlcToYaskawa.bCallMasterJob := FALSE;
	Yaskawa.stPlcToYaskawa.bExternalStart := FALSE;
	Yaskawa.stPlcToYaskawa.bExternalHold := Yaskawa.stYaskawaToPlc.bOperatingRunning
										     AND NOT Yaskawa.stYaskawaToPlc.bAlarmErrorOccured;

	etYaskawaStart := ET_YaskawaStart_eWaitExecute;              (* Next step *)

END_IF

bRunning := Yaskawa.stYaskawaToPlc.bOperatingRunning;
Yaskawa.stPlcToYaskawa.nPrgNo := nPrgNo;

(* Send command *)
CASE etYaskawaStart OF

	ET_YaskawaStart_eWaitExecute:
		bBusy := FALSE;                                     	(* Program not busy *)
		bError := FALSE;                         		(* Program not error *)

		IF rtStart.Q
     		     AND bAutoHand			(* Automatic *)
		     AND NOT bStop
		THEN
			nWatchdog := 0;
			bDone:= FALSE;                               		(* Program done *)
			bInterrupted := FALSE;				(* Program interrupted *)
			bBusy := TRUE;                                  	(* Program busy *)
			udnErrorNo := 0;                         		(* Error number *)

			wDoneFlag := 0;

			tonWatchdog(IN := FALSE);

			Yaskawa.stPlcToYaskawa.bCallMasterJob := FALSE;
			Yaskawa.stPlcToYaskawa.bExternalStart := FALSE;

			IF NOT bAutoHand
			     AND Yaskawa.stYaskawaToPlc.bHold
			THEN
				Yaskawa.stPlcToYaskawa.bExternalHold := FALSE;

				etYaskawaStart := ET_YaskawaStart_eExternalStart;              (* Next step *)
			ELSE
				Yaskawa.stPlcToYaskawa.bExternalHold := FALSE;

				etYaskawaStart := ET_YaskawaStart_eCallMasterJob;              (* Next step *)
			END_IF
		END_IF

	ET_YaskawaStart_eCallMasterJob:
		nWatchdog := nWatchdog + 1;

		Yaskawa.stPlcToYaskawa.bCallMasterJob := TRUE;

		IF Yaskawa.stYaskawaToPlc.bTopMasterJob
		     AND Yaskawa.stYaskawaToPlc.bServoIsOn
		     AND NOT Yaskawa.stYaskawaToPlc.bAlarmErrorOccured
		THEN
			nWatchdog := 0;

			Yaskawa.stPlcToYaskawa.bCallMasterJob := FALSE;

			etYaskawaStart := ET_YaskawaStart_eExternalStart;              (* Next step *)

		ELSIF Yaskawa.stYaskawaToPlc.bAlarmErrorOccured
			    OR nWatchdog > 1000
		THEN
			Yaskawa.stPlcToYaskawa.bCallMasterJob := FALSE;

			udnErrorNo := 1;                     (* Error number *)

			etYaskawaStart := ET_YaskawaStart_eError;              (* Next step *)

		END_IF

	ET_YaskawaStart_eExternalStart:
		nWatchdog := nWatchdog + 1;

		Yaskawa.stPlcToYaskawa.bExternalStart := TRUE;

		IF Yaskawa.stYaskawaToPlc.bOperatingRunning
		THEN
			wDoneFlag.0 := TRUE;
		END_IF

		IF NOT Yaskawa.stYaskawaToPlc.bPrgDone
		THEN
			wDoneFlag.1 := TRUE;
		END_IF

		IF wDoneFlag.0
		     AND wDoneFlag.1
		     AND Yaskawa.stYaskawaToPlc.bServoIsOn
		     AND NOT Yaskawa.stYaskawaToPlc.bAlarmErrorOccured
		THEN
			nWatchdog := 0;
			wDoneFlag := 0;

			Yaskawa.stPlcToYaskawa.bCallMasterJob := FALSE;
			Yaskawa.stPlcToYaskawa.bExternalStart := FALSE;

			etYaskawaStart := ET_YaskawaStart_eWfPrgDone;              (* Next step *)

		ELSIF Yaskawa.stYaskawaToPlc.bAlarmErrorOccured
			    OR nWatchdog > 1000
		THEN
			wDoneFlag := 0;

			Yaskawa.stPlcToYaskawa.bExternalStart := FALSE;

			udnErrorNo := 2;                     (* Error number *)

			etYaskawaStart := ET_YaskawaStart_eError;              (* Next step *)

		END_IF

	ET_YaskawaStart_eWfPrgDone:
		IF Yaskawa.stYaskawaToPlc.bPrgDone
	     	    AND NOT Yaskawa.stYaskawaToPlc.bAlarmErrorOccured
		THEN
			Yaskawa.stPlcToYaskawa.bCallMasterJob := FALSE;;
			Yaskawa.stPlcToYaskawa.bExternalStart := FALSE;

			etYaskawaStart := ET_YaskawaStart_eDone;              (* Next step *)

		ELSIF Yaskawa.stYaskawaToPlc.bAlarmErrorOccured
		THEN
			Yaskawa.stPlcToYaskawa.bCallMasterJob := FALSE;;
			Yaskawa.stPlcToYaskawa.bExternalStart := FALSE;

			udnErrorNo := 3;                     (* Error number *)

			etYaskawaStart := ET_YaskawaStart_eError;              (* Next step *)

		END_IF

	ET_YaskawaStart_eInterrupted:
		bInterrupted := TRUE;                                      	(* Program interrupted *)
		bBusy := FALSE;                                     		(* Program not busy *)

		etYaskawaStart := ET_YaskawaStart_eNoExecute;            		(* Next step *)

	ET_YaskawaStart_eDone:
		bDone := TRUE;						(* Command done *)
		bBusy := FALSE;						(* Command busy *)

		etYaskawaStart := ET_YaskawaStart_eNoExecute;

	ET_YaskawaStart_eError:
		bBusy := FALSE;						(* Command busy *)
		bError := TRUE;						(* Command error  *)

		etYaskawaStart := ET_YaskawaStart_eNoExecute;

	ET_YaskawaStart_eNoExecute:
		IF NOT bStart
		THEN
			(* Reset outputs *)
			bDone := FALSE;						(* Command done *)
			bInterrupted := FALSE;				(* Program interrupted *)
			bBusy := FALSE;						(* Command busy *)
			bError := FALSE;						(* Command error  *)

			nWatchdog := 0;

			etYaskawaStart := ET_YaskawaStart_eWaitExecute;
		END_IF
END_CASE;

END_FUNCTION_BLOCK

// ---- POUs/Tc2 Objects/Logger/FB_Logger.TcPOU
FUNCTION_BLOCK FB_Logger
VAR_INPUT
	bEnable								:BOOL;
	bEnableSaveInFile					:BOOL;				(* Enable save in file *)
	bInterrupt								:BOOL;
	sDateTime 							:STRING;			(* Actual date and time *)
	bDeleteAll							:BOOL;
	bLogOne							:BOOL := FALSE;		(* Log data only one time *)
	sFilePath							:STRING := 'C:\TwinCAT\Boot\';			(* Login file path *)
	sFileSuffix							:STRING := 'log';							(* Suffix of loggin file *)
	arsLogVars							:ARRAY[1..unNUM_OF_LOG_VAR] OF STRING(10);
	unLogMaxNo							:UINT;
	unLogBeforMaxNo					:UINT;
	unLogDuringMaxNo					:UINT;
	unLogAfterMaxNo						:UINT;
END_VAR
VAR_OUTPUT
	bBusy								:BOOL;
	bDone								:BOOL;
	bError								:BOOL;
	bEStop								:BOOL;
	arstLogger							:ARRAY[1..unLOG_MAX_NO] OF ST_Logger;
	arstLoggerWaitInterrupt					:ARRAY[1..unLOG_BEFOR_MAX_NO] OF ST_LoggerVar;
	arstLoggerDuringInterrupt				:ARRAY[1..unLOG_DURING_MAX_NO] OF ST_LoggerVar;
	arstLoggerAfterInterrupt					:ARRAY[1..unLOG_AFTER_MAX_NO] OF ST_LoggerVar;
END_VAR
VAR
	bFirstTime							:BOOL;
	nIdx									:INT;			(* Index *)
	udnCycleNo							:UDINT;
	unInstanceIdx							:UINT;

	unState								:UINT := 0;
	unIncLog								:UINT := 1;
	unIncDuringInterrupt					:UINT := 1;
	unIncAfterInterrupt						:UINT := 1;

	rtDeleteAll							:R_TRIG;
	rtInterrupt								:R_TRIG;
	fbLoggerFile							:FB_LoggerFile;

END_VAR
VAR CONSTANT
	unWaitInterrupt						:UINT := 0;
	unDuringInterrupt						:UINT := 1;
	unAfterInterrupt						:UINT := 2;
	unChkFile							:UINT := 3;
	unNoInterrupt							:UINT := 4;
END_VAR

IF NOT bEnable
THEN
	bBusy := FALSE;
	bDone := FALSE;
	bError := FALSE;
	bEStop := FALSE;
	bFirstTime := FALSE;
	RETURN;
END_IF

IF NOT bFirstTime
THEN
	bBusy := FALSE;
	bDone := FALSE;
	bError := FALSE;
	bEStop := FALSE;
	unState := 0;
	unIncLog := 1;
	unIncDuringInterrupt := 1;
	unIncAfterInterrupt := 1;

	unLOG_INSTANCE_IDX  := unLOG_INSTANCE_IDX + 1;
	unInstanceIdx := unLOG_INSTANCE_IDX;

	unState := unWaitInterrupt;

	bFirstTime := TRUE;
END_IF


rtDeleteAll(CLK := bDeleteAll);

IF rtDeleteAll.Q
    AND (bDone OR bError)
THEN
	bBusy := FALSE;
	bDone := FALSE;
	bError := FALSE;
	bEStop := FALSE;
	unState := 0;
	unIncLog := 1;
	unIncDuringInterrupt := 1;
	unIncAfterInterrupt := 1;

	unState := unWaitInterrupt;
END_IF

rtInterrupt(CLK := bInterrupt);
IF rtInterrupt.Q
THEN
	unState := unWaitInterrupt;
END_IF;

udnCycleNo := udnCycleNo + 1;

CASE unState OF
	
	unWaitInterrupt:
		bBusy := FALSE;
		bDone := FALSE;
		bError := FALSE;

		fbLoggerFile.bExecute := FALSE;

		(* Shift down logger list by 1 *)
		A_ShiftDown();

		(* Write time stamp and value of variables before interrupt *)
		arstLoggerWaitInterrupt[1].udnCycleNo := udnCycleNo;
		arstLoggerWaitInterrupt[1].sTimeStamp := sDateTime;
		arstLoggerWaitInterrupt[1].arsLogVars := arsLogVars;

		IF bInterrupt
		THEN
			bBusy := TRUE;
			bDone := FALSE;

			bEStop := bLogOne;

			MEMSET(ADR(arstLoggerDuringInterrupt), 0, SIZEOF(arstLoggerDuringInterrupt));
			MEMSET(ADR(arstLoggerAfterInterrupt), 0, SIZEOF(arstLoggerAfterInterrupt));

			(* Log data *)
			IF unIncLog <= unLOG_MAX_NO
			THEN
				MEMCPY(ADR(arstLogger[unIncLog].arstLoggerWaitInterrupt), ADR(arstLoggerWaitInterrupt), SIZEOF(arstLoggerWaitInterrupt));
			ELSE
				unIncLog := 1;
				MEMCPY(ADR(arstLogger[unIncLog].arstLoggerWaitInterrupt), ADR(arstLoggerWaitInterrupt), SIZEOF(arstLoggerWaitInterrupt));
			END_IF

			(* Write time stamp and value of variables during interrupt *)
			unIncDuringInterrupt := 1;
			arstLoggerDuringInterrupt[unIncDuringInterrupt].udnCycleNo := udnCycleNo;
			arstLoggerDuringInterrupt[unIncDuringInterrupt].sTimeStamp := sDateTime;
			arstLoggerDuringInterrupt[unIncDuringInterrupt].arsLogVars := arsLogVars;
			unIncDuringInterrupt := unIncDuringInterrupt + 1;

			fbLoggerFile.sFileName := CONCAT(
										sDateTime,
										CONCAT(
											'_',
											UINT_TO_STRING(unInstanceIdx)
										)
									);

			unState := unDuringInterrupt;

		END_IF

	unDuringInterrupt:
		IF unIncDuringInterrupt <= unLOG_DURING_MAX_NO
		THEN
			(*  Write time stamp and value of variables during interrupt *)
			arstLoggerDuringInterrupt[unIncDuringInterrupt].udnCycleNo := udnCycleNo;
			arstLoggerDuringInterrupt[unIncDuringInterrupt].sTimeStamp := sDateTime;
			arstLoggerDuringInterrupt[unIncDuringInterrupt].arsLogVars := arsLogVars;
		
			unIncDuringInterrupt := unIncDuringInterrupt + 1;

		END_IF

		IF NOT bInterrupt
		THEN
			(* Log data *)
			MEMCPY(ADR(arstLogger[unIncLog].arstLoggerDuringInterrupt), ADR(arstLoggerDuringInterrupt), SIZEOF(arstLoggerDuringInterrupt));

			(* Write time stamp and value of variables after interrupt *)
			unIncAfterInterrupt := 1;
			arstLoggerAfterInterrupt[unIncAfterInterrupt].udnCycleNo := udnCycleNo;
			arstLoggerAfterInterrupt[unIncAfterInterrupt].sTimeStamp := sDateTime;
			arstLoggerAfterInterrupt[unIncAfterInterrupt].arsLogVars := arsLogVars;
			unIncAfterInterrupt := unIncAfterInterrupt + 1;

			unState := unAfterInterrupt;

		END_IF

	unAfterInterrupt:
		IF unIncAfterInterrupt <= unLOG_AFTER_MAX_NO
		THEN
			(* Write time stamp and value of variables after interrupt *)
			arstLoggerAfterInterrupt[unIncAfterInterrupt].udnCycleNo := udnCycleNo;
			arstLoggerAfterInterrupt[unIncAfterInterrupt].sTimeStamp := sDateTime;	
			arstLoggerAfterInterrupt[unIncAfterInterrupt].arsLogVars := arsLogVars;

			unIncAfterInterrupt := unIncAfterInterrupt + 1;
		ELSE
			(* Log data *)
			MEMCPY(ADR(arstLogger[unIncLog].arstLoggerAfterInterrupt), ADR(arstLoggerAfterInterrupt), SIZEOF(arstLoggerAfterInterrupt));

			fbLoggerFile.bExecute := TRUE;

			IF fbLoggerFile.bBusy
			THEN
				unState := unChkFile;

			ELSIF fbLoggerFile.bError
			THEN
				fbLoggerFile.bExecute := FALSE;
	
				bBusy := FALSE;
				bError := TRUE;
	
				unState := unNoInterrupt;

			END_IF
		END_IF

	unChkFile:
		IF NOT bEnableSaveInFile
		     OR fbLoggerFile.bDone
		THEN
			fbLoggerFile.bExecute := FALSE;

			bBusy := FALSE;
			bDone := TRUE;

			unState := unNoInterrupt;

		ELSIF  fbLoggerFile.bError
		THEN
			fbLoggerFile.bExecute := FALSE;

			bBusy := FALSE;
			bError := TRUE;

			unState := unNoInterrupt;

		END_IF

	unNoInterrupt:
		IF NOT bInterrupt
		    AND NOT bEStop
		THEN
			bBusy := FALSE;
			bDone := FALSE;
			bError := FALSE;

			unIncLog := unIncLog + 1;

			unState := unWaitInterrupt;
		END_IF

END_CASE


fbLoggerFile(
	bEnable := bEnableSaveInFile,
	sFilePath := sFilePath,
	sFileSuffix := sFileSuffix,
	arstLoggerWaitInterrupt := arstLoggerWaitInterrupt,
	arstLoggerDuringInterrupt := arstLoggerDuringInterrupt,
	arstLoggerAfterInterrupt := arstLoggerAfterInterrupt
 );

ACTION A_ShiftDown:

FOR nIdx := unLOG_BEFOR_MAX_NO - 1 TO 1 BY -1
DO
	arstLoggerWaitInterrupt[nIdx + 1] := arstLoggerWaitInterrupt[nIdx];
END_FOR
END_ACTION

END_FUNCTION_BLOCK

// ---- POUs/Tc2 Objects/Logger/FB_LoggerFile.TcPOU
FUNCTION_BLOCK FB_LoggerFile
(*

This function block is used to write loggin datas into file.

Constructor: 		Patryk Panylo
Company:		E. Riexinger GmbH
Date:			25.03.2014
Version:			1.00

Date:			Revision:		Who:				Comment
dd.mm.yyyy		x.xx			Initials			comment

*)

VAR_INPUT
	bEnable						:BOOL;					(* Enable FB *)
	bExecute					:BOOL;					(* Execute operation *)
	sFilePath					:STRING;				(* File path *)
	sFileName					:STRING;				(* File name *)
	sFileSuffix					:STRING := 'dat';			(* Suffix of file *)
	arstLoggerWaitInterrupt			:ARRAY[1..unLOG_BEFOR_MAX_NO] OF ST_LoggerVar;			(* Data to write to file *)
	arstLoggerDuringInterrupt		:ARRAY[1..unLOG_DURING_MAX_NO] OF ST_LoggerVar;			(* Data to write to file *)
	arstLoggerAfterInterrupt			:ARRAY[1..unLOG_AFTER_MAX_NO] OF ST_LoggerVar;			(* Data to write to file *)
	tTimeout						:TIME := t#1s;				(* States the time before the function is cancelled *)
END_VAR
VAR_OUTPUT
	bBusy						:BOOL;					(* Program busy *)
	bDone						:BOOL;					(* Program done *)
	bError						:BOOL;					(* Program error *)
	udnErrNo					:UDINT;					(* Error number *)
END_VAR
VAR_IN_OUT

END_VAR
VAR
	(* Enummerations *)
	enStep						: (eWaitExecute := 0, eChkFileName, eChkeNumOfRecords, eFileOpen, eChkFileOpen, eFilePuts, eChkFilePuts, eFileClose, eChkFileClose, eDone, eError, eNotExecute);			(* Sequence state for open, read/write and close the file *)
	enGetData					: (eWaitInterruptData, eDuringInterruptData, eAfterInterruptData, eNoData);					(* Sequence state for data *)

	(* Variables *)
	bFirstTime					:BOOL;					(* First PLC cycle *)
	unLogSize					:UINT;
	unLogIdx						:UINT;
	unRecordsSize				:UINT;
	unRecordsIdx					:UINT;

	dwMode						:DWORD;				(* Contains the mode in which the file is to be opened *)
	sPathName					:STRING;				(* Contains the path and filename for the file to be opened *)
	hFileHandle					:UINT;					(* File handle *)

	unPutsCounter				:UINT;

	sRecordsToWrite				:STRING;

	(* Instances *)
	fbFileOpen					:FB_FileOpen;			(* File open *)
	fbFileClose					:FB_FileClose;			(* File close *)
	fbFilePuts					:FB_FilePuts;				(* File puts *)

END_VAR
VAR CONSTANT
	sSeparator					:STRING := '$T';
	sNewLine					:STRING := '$N'; 							(* End line sign for lines *)
END_VAR

IF NOT bEnable				(* Enable FB *)
THEN
	bFirstTime := FALSE;		(* First PLC cycle *)
	bBusy := FALSE;			(* Program busy *)
	bDone := FALSE;			(* Program done *)
	bError := FALSE;			(* Program error *)
	udnErrNo := 0;				(* Error number *)
	RETURN;
END_IF

IF NOT bFirstTime
THEN
	bBusy := FALSE;			(* Program busy *)
	bDone := FALSE;			(* Program done *)
	bError := FALSE;			(* Program error *)

	enStep := eWaitExecute;

	bFirstTime := TRUE;
END_IF


(* Sequence state for open, read/write and close the file *)
CASE enStep
OF

	eWaitExecute:
		IF bExecute
		THEN
			fbFileOpen.bExecute := FALSE;			(* File open *)
			fbFileClose.bExecute := FALSE;			(* File close *)
			fbFilePuts.bExecute := FALSE;			(* File puts *)

			bBusy := TRUE;
			bDone := FALSE;
			bError := FALSE;
			udnErrNo := 0;

			dwMode := FOPEN_MODEWRITE OR FOPEN_MODETEXT;

			enStep := eChkFileName;			(* Next step *)

		END_IF

	(* Check file name and path *)
	eChkFileName:

		sPathName := CONCAT(
						sFilePath, CONCAT(
									sFileName, CONCAT(
												'.', sFileSuffix)));

		IF sFilePath <> ''
		     AND sFileName <> ''
		     AND sFileSuffix <> ''
		THEN
			enStep := eChkeNumOfRecords;			(* Next step *)

		ELSE
			udnErrNo := eChkFileName;

			enStep := eError;				(* Next step *)

		END_IF

	(* Check number of records to save *)
	eChkeNumOfRecords:
		IF unNUM_OF_LOG_VAR = 0
		THEN
			enStep := eDone;				(* Next step *)
	
		ELSE
			enStep := eFileOpen;			(* Next step *)

		END_IF
	(* Open the file *)
	eFileOpen:
		fbFileOpen.bExecute := TRUE;

		enStep := eChkFileOpen;				(* Next step *)

	(* Check open the file *)
	eChkFileOpen:
		IF NOT fbFileOpen.bBusy
		THEN
			IF NOT fbFileOpen.bError
			THEN
				fbFileOpen.bExecute := FALSE;
				hFileHandle := fbFileOpen.hFile;

				unLogIdx := 0;
		  		unRecordsIdx := 0;

				enGetData := eWaitInterruptData;
				enStep := eFilePuts;			(* Next step *)

			ELSE
				fbFileOpen.bExecute := FALSE;
				udnErrNo := fbFileOpen.nErrId;
	
				enStep := eError;					(* Next step *)

			END_IF
		END_IF

	(* Puts data into the file *)
	eFilePuts:
		(* Get data *)
		A_GetData();

		IF LEN(sRecordsToWrite) > 254
		THEN
			sRecordsToWrite := DELETE(
								sRecordsToWrite,
								LEN(sRecordsToWrite) + 1 - 254, 254
							    );
		END_IF


		sRecordsToWrite := CONCAT(
							sRecordsToWrite,
							SEL(unRecordsIdx = 0, sSeparator, sNewLine)
						    );


		fbFilePuts.bExecute := TRUE;

		enStep := eChkFilePuts;				(* Next step *)

	(* Check puts the file *)
	eChkFilePuts:
		IF NOT fbFilePuts.bBusy
		THEN
			IF NOT fbFilePuts.bError
			THEN
				fbFilePuts.bExecute := FALSE;
				unPutsCounter := unPutsCounter + 1;

				IF enGetData = eNoData
				THEN
					enStep := eFileClose;				(* Next step *)
				ELSE
					enStep := eFilePuts;				(* Next step *)
				END_IF

			ELSIF  fbFilePuts.bError
			THEN
				fbFilePuts.bExecute := FALSE;
				udnErrNo := fbFilePuts.nErrId;

				enStep := eError;					(* Next step *)

			END_IF
		END_IF

	(* Close the file *)
	eFileClose:
		fbFileClose.bExecute := TRUE;

		enStep := eChkFileClose;				(* Next step *)

	(* Check close the file *)
	eChkFileClose:
		IF NOT fbFileClose.bBusy
		THEN
			IF NOT fbFileClose.bError
			THEN
				fbFileClose.bExecute := FALSE;
				enStep := eDone;					(* Next step *)

				IF bError
				THEN
					enStep := eError;				(* Next step *)
				END_IF

			ELSE
				fbFileClose.bExecute := FALSE;
				udnErrNo := fbFileClose.nErrId;
	
				enStep := eError;					(* Next step *)
				
			END_IF
		END_IF

	eDone:
		bBusy := FALSE;
		bDone := TRUE;
		bError := FALSE;
		udnErrNo := 0;

		enStep := eNotExecute;					(* Next step *)

	eError:
		IF NOT bError
		     AND hFileHandle <> 0
		THEN
			bDone := FALSE;
			bError := TRUE;

			enStep := eFileClose;					(* Next step *)

		ELSE
			bBusy := FALSE;
			bDone := FALSE;
			bError := TRUE;
	
			enStep := eNotExecute;					(* Next step *)
		END_IF

	eNotExecute:
		IF NOT bExecute
		THEN
			bBusy := FALSE;
			bDone := FALSE;
			bError := FALSE;
			udnErrNo := 0;

			enStep := eWaitExecute;			(* Next step *)

		END_IF

END_CASE

fbFileOpen(
	sNetId := '',
	sPathName := sPathName,
	nMode := dwMode,
	ePath := PATH_GENERIC,
	tTimeout := tTimeout
);
fbFileClose(
	sNetId := '',
	hFile := hFileHandle,
	tTimeout := tTimeout
);
fbFilePuts(
	sNetId := '',
	hFile:= hFileHandle,
	sLine := sRecordsToWrite,
	tTimeout := tTimeout
 );

ACTION A_GetData:

CASE enGetData
OF
	eWaitInterruptData:
		IF unLogIdx = 0
		THEN
			unLogIdx := 1;
			unLogSize := unLOG_BEFOR_MAX_NO;

			sRecordsToWrite := '[WAIT INTERRUPT]';

		ELSIF unRecordsIdx = 0
		THEN
			unRecordsIdx	 := 1;
			unRecordsSize := unNUM_OF_LOG_VAR;

			sRecordsToWrite := CONCAT(
								UDINT_TO_STRING(arstLoggerWaitInterrupt[unLogIdx].udnCycleNo),
								CONCAT(
									sSeparator,
									arstLoggerWaitInterrupt[unLogIdx].sTimeStamp
								)
							   );

		ELSE

			sRecordsToWrite := arstLoggerWaitInterrupt[unLogIdx].arsLogVars[unRecordsIdx];

			unRecordsIdx := unRecordsIdx + 1;

			IF unRecordsIdx > unRecordsSize
			THEN
				unRecordsIdx := 0;
				unLogIdx := unLogIdx + 1;
			END_IF

		END_IF

		IF unLogIdx > unLogSize
		THEN
			unLogIdx := 0;
		  	unRecordsIdx := 0;
			enGetData := eDuringInterruptData;					(* Next step *)
		END_IF

	eDuringInterruptData:

		IF unLogIdx = 0
		THEN
			unLogIdx := 1;
			unLogSize := unLOG_DURING_MAX_NO;

			sRecordsToWrite := '[DURING INTERRUPT]';

		ELSIF unRecordsIdx = 0
		THEN
			unRecordsIdx	 := 1;
			unRecordsSize := unNUM_OF_LOG_VAR;

			sRecordsToWrite := CONCAT(
								UDINT_TO_STRING(arstLoggerDuringInterrupt[unLogIdx].udnCycleNo),
								CONCAT(
									sSeparator,
									arstLoggerDuringInterrupt[unLogIdx].sTimeStamp
								)
							   );

		ELSE
			sRecordsToWrite := arstLoggerDuringInterrupt[unLogIdx].arsLogVars[unRecordsIdx];

			unRecordsIdx := unRecordsIdx + 1;

			IF unRecordsIdx > unRecordsSize
			THEN
				unRecordsIdx := 0;
				unLogIdx := unLogIdx + 1;
			END_IF

		END_IF

		IF unLogIdx > unLogSize
		THEN
			unLogIdx := 0;
		  	unRecordsIdx := 0;
			enGetData := eAfterInterruptData;					(* Next step *)
		END_IF

	eAfterInterruptData:

		IF unLogIdx = 0
		THEN
			unLogIdx := 1;
			unLogSize := unLOG_AFTER_MAX_NO;

			sRecordsToWrite := '[AFTER INTERRUPT]';

			IF LEN(arstLoggerAfterInterrupt[unLogIdx].sTimeStamp) = 0
			THEN
				unLogIdx := unLOG_AFTER_MAX_NO + 1;
			END_IF

		ELSIF unRecordsIdx = 0
		THEN
			unRecordsIdx	 := 1;
			unRecordsSize := unNUM_OF_LOG_VAR;

			sRecordsToWrite := CONCAT(
								UDINT_TO_STRING(arstLoggerAfterInterrupt[unLogIdx].udnCycleNo),
								CONCAT(
									sSeparator,
									arstLoggerAfterInterrupt[unLogIdx].sTimeStamp
								)
							   );

		ELSE
			sRecordsToWrite := arstLoggerAfterInterrupt[unLogIdx].arsLogVars[unRecordsIdx];

			unRecordsIdx := unRecordsIdx + 1;

			IF unRecordsIdx > unRecordsSize
			THEN
				unRecordsIdx := 0;
				unLogIdx := unLogIdx + 1;
			END_IF

		END_IF

		IF unLogIdx > unLogSize
		THEN
			unLogIdx := 0;
		  	unRecordsIdx := 0;
			enGetData := eNoData;
		END_IF

	eNoData:
		unLogIdx := 0;
		 unRecordsIdx := 0;

END_CASE
END_ACTION

END_FUNCTION_BLOCK

// ---- POUs/Tc2 Objects/Logic/F_DwordToBitReal.TcPOU
FUNCTION F_DwordToBitReal : REAL
VAR_INPUT
	dwIn : DWORD;
END_VAR
VAR
	pt : POINTER TO REAL;
END_VAR

pt := ADR(dwIn);
F_DwordToBitReal := pt^;

END_FUNCTION

// ---- POUs/Tc2 Objects/Logic/F_RealToBitDword.TcPOU
FUNCTION F_RealToBitDword : DWORD
VAR_INPUT
	rIn : REAL;
END_VAR
VAR
	pt : POINTER TO DWORD;
END_VAR

pt := ADR(rIn);
F_RealToBitDword := pt^;

END_FUNCTION

// ---- POUs/Tc2 Objects/Logic/F_ResetBitOfDWord.TcPOU
FUNCTION F_ResetBitOfDWord : DWORD
VAR_INPUT
	dwInput			:DWORD;
	usnBitNr			:USINT;
END_VAR
VAR
END_VAR

F_ResetBitOfDWord := dwInput;
CASE usnBitNr OF
	0:
	F_ResetBitOfDWord.0 := FALSE;
	1:
	F_ResetBitOfDWord.1 := FALSE;
	2:
	F_ResetBitOfDWord.2 := FALSE;
	3:
	F_ResetBitOfDWord.3 := FALSE;
	4:
	F_ResetBitOfDWord.4 := FALSE;
	5:
	F_ResetBitOfDWord.5 := FALSE;
	6:
	F_ResetBitOfDWord.6 := FALSE;
	7:
	F_ResetBitOfDWord.7 := FALSE;
	8:
	F_ResetBitOfDWord.8 := FALSE;
	9:
	F_ResetBitOfDWord.9 := FALSE;
	10:
	F_ResetBitOfDWord.10 := FALSE;
	11:
	F_ResetBitOfDWord.11 := FALSE;
	12:
	F_ResetBitOfDWord.12 := FALSE;
	13:
	F_ResetBitOfDWord.13 := FALSE;
	14:
	F_ResetBitOfDWord.14 := FALSE;
	15:
	F_ResetBitOfDWord.15 := FALSE;
	16:
	F_ResetBitOfDWord.16 := FALSE;
	17:
	F_ResetBitOfDWord.17 := FALSE;
	18:
	F_ResetBitOfDWord.18 := FALSE;
	19:
	F_ResetBitOfDWord.19 := FALSE;
	20:
	F_ResetBitOfDWord.20 := FALSE;
	21:
	F_ResetBitOfDWord.21 := FALSE;
	22:
	F_ResetBitOfDWord.22 := FALSE;
	23:
	F_ResetBitOfDWord.23 := FALSE;
	24:
	F_ResetBitOfDWord.24 := FALSE;
	25:
	F_ResetBitOfDWord.25 := FALSE;
	26:
	F_ResetBitOfDWord.26 := FALSE;
	27:
	F_ResetBitOfDWord.27 := FALSE;
	28:
	F_ResetBitOfDWord.28 := FALSE;
	29:
	F_ResetBitOfDWord.29 := FALSE;
	30:
	F_ResetBitOfDWord.30 := FALSE;
	31:
	F_ResetBitOfDWord.31 := FALSE;
END_CASE

END_FUNCTION

// ---- POUs/Tc2 Objects/Logic/F_SetBitOfDWord.TcPOU
FUNCTION F_SetBitOfDWord : DWORD
VAR_INPUT
	dwInput			:DWORD;
	usnBitNr			:USINT;
END_VAR
VAR
END_VAR

F_SetBitOfDWord := dwInput;
CASE usnBitNr OF
	0:
	F_SetBitOfDWord.0 := TRUE;
	1:
	F_SetBitOfDWord.1 := TRUE;
	2:
	F_SetBitOfDWord.2 := TRUE;
	3:
	F_SetBitOfDWord.3 := TRUE;
	4:
	F_SetBitOfDWord.4 := TRUE;
	5:
	F_SetBitOfDWord.5 := TRUE;
	6:
	F_SetBitOfDWord.6 := TRUE;
	7:
	F_SetBitOfDWord.7 := TRUE;
	8:
	F_SetBitOfDWord.8 := TRUE;
	9:
	F_SetBitOfDWord.9 := TRUE;
	10:
	F_SetBitOfDWord.10 := TRUE;
	11:
	F_SetBitOfDWord.11 := TRUE;
	12:
	F_SetBitOfDWord.12 := TRUE;
	13:
	F_SetBitOfDWord.13 := TRUE;
	14:
	F_SetBitOfDWord.14 := TRUE;
	15:
	F_SetBitOfDWord.15 := TRUE;
	16:
	F_SetBitOfDWord.16 := TRUE;
	17:
	F_SetBitOfDWord.17 := TRUE;
	18:
	F_SetBitOfDWord.18 := TRUE;
	19:
	F_SetBitOfDWord.19 := TRUE;
	20:
	F_SetBitOfDWord.20 := TRUE;
	21:
	F_SetBitOfDWord.21 := TRUE;
	22:
	F_SetBitOfDWord.22 := TRUE;
	23:
	F_SetBitOfDWord.23 := TRUE;
	24:
	F_SetBitOfDWord.24 := TRUE;
	25:
	F_SetBitOfDWord.25 := TRUE;
	26:
	F_SetBitOfDWord.26 := TRUE;
	27:
	F_SetBitOfDWord.27 := TRUE;
	28:
	F_SetBitOfDWord.28 := TRUE;
	29:
	F_SetBitOfDWord.29 := TRUE;
	30:
	F_SetBitOfDWord.30 := TRUE;
	31:
	F_SetBitOfDWord.31 := TRUE;
END_CASE

END_FUNCTION

// ---- POUs/Tc2 Objects/MachineEquipment/F_kFeedReductionSlowGuidings.TcPOU
FUNCTION F_kFeedReductionSlowGuidings : LREAL
(*

The function used to reduction saw feed dependent of slow sawband guidings 
Output factor: 0..1 (1=no speed reduction)

Constructor: 		Eduard Schüle
Company:		E. Riexinger GmbH
Date:			20.11.2015
Version:			1.01

Date:		Revision:	Who:	Comment
24.11.2015	1.01			ES		speed reduction only if for guidings required

*)
VAR_INPUT
	(* Input variables / Eingang Variablen *)
	bEnable							:BOOL;						(* Function block enable *)
	lrActPos							:LREAL;						(* Current position of axis *)
	lrActSawbowAngle				:LREAL;						(* SawBow Angle, cutting angle *)
	lrActGuiding1Position				:LREAL;
	lrActGuiding2Position				:LREAL;
	lrVerticalOffset					:LREAL;						(* vertical offset collision contour *)
	lrActSpeed						:LREAL;						(* Current speed of axis *)
	lrActVelo							:LREAL;						(* Current Velocity for axis *)
	lrMaxVelo						:LREAL;						(* Max Velocity of axis *)
	lrMaxMaster						:LREAL;						(* max. Velocity Master *)
	lrMaxSlave						:LREAL;						(* max. Velocity Slave *)
	lrMinK							:LREAL;						(* minimum Speedfactor, 0.0 .. 1.0 *)
	lrCStartMaxPos					:LREAL;						(* Contour start maximal position *)
	lrCEndMinPos					:LREAL;						(* Contour end minimal position  *)
	lrCSafetyDistance					:LREAL;						(* Safety distance *)
	lrTableHeight						:LREAL;						(* Table height, if need guidings go to table width *)
	lrTableWidth						:LREAL;						(* table width *)
	lrGuidingMinPos					:LREAL;						(* sawband guiding min position, below no speed reduction *)
	lrGuidingMaxPos					:LREAL;						(* sawband guiding max position, above no speed reduction *)
	lrGuidingWindow					:LREAL;						(* sawband guiding position window *)
END_VAR
VAR
	(* Variables *)
	lrActPosCache					:LREAL;						(* intern position of axis *)
	lrCRadius						:LREAL;						(* Radius *)
	lrCMiddlePos						:LREAL;						(* Middle position *)
	lrCAlfa							:LREAL;						(* Angle of inclination *)
	lrTanAlfa							:LREAL;						(* Tangent of alfa *)
	lrAngleFactor						:LREAL;						(* Sawbow angle factor, ellipse *)
	lrSpeedFactor					:LREAL;						(*  *)
	lrVelo							:LREAL;						(*  *)
	lrCStartMaxPosCache 				:LREAL;
	lrCEndMinPosCache 				:LREAL;
	lrActGuidingSetPosition			:LREAL;
	lrActPosN1						:LREAL;						(*  position of axis last cycle *)
END_VAR

IF NOT bEnable
THEN
	F_kFeedReductionSlowGuidings := lrActVelo;
	RETURN;
END_IF

lrActGuidingSetPosition := F_CalcContour(
	etContourType := ET_ContourType_eEllipse,
	lrActPos := lrActPos,
	lrActAngle := lrActSawbowAngle,
	lrVerticalOffset := lrVerticalOffset,
	lrStartMaxPos := lrCStartMaxPos,
	lrEndMinPos := lrCEndMinPos,
	lrSafetyDistance := lrCSafetyDistance-20.0,
	lrTableHeight := lrTableHeight,
	lrTableWidth := lrTableWidth,
	lrActVeloExt := 0
	);

lrCStartMaxPosCache := lrCStartMaxPos + ABS(lrCSafetyDistance + 50.0);
lrCEndMinPosCache := lrCEndMinPos - ABS(lrCSafetyDistance + 50.0);

lrCRadius := ABS(lrCStartMaxPosCache - lrCEndMinPos) / 2;
lrCMiddlePos := lrCEndMinPosCache + lrCRadius;										(* Middle position *)

lrActPosCache := lrActPos - lrVerticalOffset;

IF lrActPos >= lrTableHeight
THEN
	IF (lrActPosCache <= lrCStartMaxPosCache)
		AND (lrActPosCache >= lrCEndMinPosCache)
		AND lrCRadius > 0.0
(*		AND NOT(lrActGuiding1Position < (lrGuidingMinPos + lrGuidingWindow)) (* nicht wenn MIN Position *)
		AND NOT(lrActGuiding2Position < (lrGuidingMinPos + lrGuidingWindow))
		AND NOT(lrActGuiding1Position > (lrGuidingMaxPos - lrGuidingWindow))	(* not if MAX position *)
		AND NOT(lrActGuiding2Position > (lrGuidingMaxPos - lrGuidingWindow))*)
		AND NOT(lrActGuiding1Position > lrActGuidingSetPosition)
		AND NOT(lrActGuiding2Position > lrActGuidingSetPosition)
(*		AND lrActSpeed < 0
		(*AND (lrActPos - lrActPosN1) < 0 (* down < 0 *)*)
		AND lrActPos > lrCMiddlePos*)
	THEN
		lrCAlfa := ACOS(ABS(lrCMiddlePos - lrActPosCache) /  lrCRadius);							(* Angle of inclination *)
		lrTanAlfa := TAN(lrCAlfa);														(* Tangent of alfa *)
		lrAngleFactor := 1 / COS( MIN(ABS(lrActSawbowAngle), 89.9) / 180.0*PI);			(* Sawbow angle factor, ellipse *)
		lrSpeedFactor := MAX(lrMinK, lrTanAlfa * lrAngleFactor);

		lrVelo := LIMIT(0, lrSpeedFactor * lrMaxSlave / lrMaxMaster * lrMaxVelo, lrMaxVelo);
	
		F_kFeedReductionSlowGuidings := MIN(lrVelo, ABS(lrActVelo));

		IF lrActVelo<0 THEN
			F_kFeedReductionSlowGuidings := -F_kFeedReductionSlowGuidings;
		END_IF

	ELSE

		F_kFeedReductionSlowGuidings := lrActVelo;

	END_IF
ELSE
	IF		 lrActGuiding1Position > (lrTableWidth / 2 + 10.0)
		AND lrActGuiding2Position > (lrTableWidth / 2 +10.0)
	THEN
		F_kFeedReductionSlowGuidings := lrActVelo;
	ELSE
		F_kFeedReductionSlowGuidings := 0;
	END_IF
END_IF

lrActPosN1 := lrActPos;

END_FUNCTION

// ---- POUs/Tc2 Objects/Mathematical/Delay/FB_Delay.TcPOU
FUNCTION_BLOCK FB_Delay
(*
Function block used to caculate delay

Constructor: 		Patryk Panylo
Company:		E. Riexinger GmbH
Date:			14.07.2014
Version:			1.00

Date:			Revision:		Who:				Comment
dd.mm.yyyy		x.xx			Initials			comment

*)
VAR_INPUT
	(* Enummerations *)

	(* Variables *)
	bEnable								:BOOL := TRUE;					(* Enable FB *)

	lrInSignal								:LREAL;							(* Input signal *)
	tDeadTime							:TIME := t#200ms;					(* Dead time *)
	tTaskCycle							:TIME := t#2ms; 					(* Cycle time *)

	(* References *)

	(* Interfaces *)

	(* Instances *)
END_VAR
VAR_OUTPUT
	(* Enummerations *)
	
	(* Variables *)
	lrOutSignal							:LREAL;							(* Output signal *)

	(* References *)

	(* Interfaces *)

	(* Instances *)
END_VAR
VAR
	(* Enummerations *)

	(* Variables *)
	bFirstTime							:BOOL;							(* First cycle *)

	lrTimeRatio							:LREAL;
	lrLastSignal							:LREAL;							(* Last signal *)

	(* References *)

	(* Interfaces *)

	(* Instances *)
	tpClock								:TP;

END_VAR

IF NOT bEnable
THEN
	lrOutSignal := lrInSignal;

	bFirstTime := FALSE;
	RETURN;
END_IF

IF NOT bFirstTime
THEN
	lrOutSignal := lrInSignal;

	tpClock(
		IN := FALSE,
		PT := tTaskCycle
	);

	bFirstTime := TRUE;
END_IF


tpClock();

IF NOT tpClock.Q
THEN
	tpClock(IN := FALSE);

	IF tDeadTime > t#0ms
	THEN
		lrTimeRatio := TIME_TO_LREAL(tTaskCycle) / TIME_TO_LREAL(tDeadTime);

		lrOutSignal := lrLastSignal + (lrInSignal - lrLastSignal) * lrTimeRatio;
	ELSE
		lrOutSignal := lrLastSignal;
	END_IF

	tpClock(IN := TRUE);
END_IF

lrLastSignal := lrOutSignal;

END_FUNCTION_BLOCK

// ---- POUs/Tc2 Objects/Mathematical/FB_Differential.TcPOU
FUNCTION_BLOCK FB_Differential
(*
Function block used to calculate differential

Constructor: 		Patryk Panylo
Company:		E. Riexinger GmbH
Date:			05.06.2014
Version:			1.00

Date:			Revision:		Who:				Comment
dd.mm.yyyy		x.xx			Initials			comment

*)
VAR_INPUT
	(* Enummerations *)
	
	(* Variables *)
	bEnable								:BOOL := TRUE;					(* Enable FB *)

	lrInSignal								:LREAL;							(* Input signal *)
	lrDifferentialValue						:LREAL := 1.0;						(* Differential value *)
	lrTaskCycle							:LREAL := 1.0; 					(* Cycle time *)

	(* References *)

	(* Interfaces *)

	(* Instances *)
END_VAR
VAR_OUTPUT
	(* Enummerations *)
	
	(* Variables *)
	lrOutSignal							:LREAL;							(* Output signal *)

	(* References *)

	(* Interfaces *)

	(* Instances *)
END_VAR
VAR
	(* Enummerations *)
	
	(* Variables *)
	bFirstTime							:BOOL;							(* First cycle *)

	lrLastSignal							:LREAL;							(* Last signal *)

	(* References *)

	(* Interfaces *)

	(* Instances *)


END_VAR

IF NOT bEnable
THEN
	lrOutSignal := lrInSignal;

	bFirstTime := FALSE;
	RETURN;
END_IF

IF NOT bFirstTime
THEN
	lrLastSignal := lrInSignal;
	bFirstTime := TRUE;
END_IF

IF lrTaskCycle > 0.0
THEN
	lrOutSignal := lrDifferentialValue * (lrInSignal - lrLastSignal) / lrTaskCycle;
ELSE
	lrOutSignal := 0.0;
END_IF
lrLastSignal := lrInSignal;

END_FUNCTION_BLOCK

// ---- POUs/Tc2 Objects/Mathematical/FB_Integral.TcPOU
FUNCTION_BLOCK FB_Integral
(*
Function block used to calculate integral

Constructor: 		Patryk Panylo
Company:		E. Riexinger GmbH
Date:			05.06.2014
Version:			1.00

Date:			Revision:		Who:				Comment
dd.mm.yyyy		x.xx			Initials			comment

*)
VAR_INPUT
	(* Enummerations *)

	(* Variables *)
	bEnable								:BOOL := TRUE;					(* Enable FB *)

	lrInSignal								:LREAL;							(* Input signal *)
	lrIntegralValue						:LREAL := 1.0;						(* Integration value in 1/sec *)
	lrTaskCycle							:LREAL := 1.0; 					(* Cycle time *)

	(* References *)

	(* Interfaces *)

	(* Instances *)
END_VAR
VAR_OUTPUT
END_VAR
VAR_IN_OUT
	(* Enummerations *)
	
	(* Variables *)
	lrOutSignal							:LREAL;							(* Output signal *)

	(* References *)

	(* Interfaces *)

	(* Instances *)
END_VAR
VAR
	(* Enummerations *)
	
	(* Variables *)
	bFirstTime							:BOOL;							(* First cycle *)

	lrLastSignal							:LREAL;							(* Last signal *)

	(* References *)

	(* Interfaces *)

	(* Instances *)


END_VAR

IF NOT bEnable
THEN
	bFirstTime := FALSE;
	RETURN;
END_IF

IF NOT bFirstTime
THEN
	lrLastSignal := lrInSignal;
	bFirstTime := TRUE;
END_IF

lrOutSignal := lrIntegralValue * lrTaskCycle * (lrInSignal + lrLastSignal) * 0.5 + lrOutSignal;
lrLastSignal := lrInSignal;

END_FUNCTION_BLOCK

// ---- POUs/Tc2 Objects/Mathematical/F_Exp10.TcPOU
FUNCTION F_Exp10 : REAL
VAR_INPUT
	X : REAL;
END_VAR


(*
version 1.0	 2 dec 2007
programmer 	hugo
tested by		tobias

this function calculates the exponent to the basis 10
exp10(3) = 1000

*)

F_Exp10 := EXP(X * 2.30258509299405);

END_FUNCTION

// ---- POUs/Tc2 Objects/Mathematical/F_FloorDN.TcPOU
FUNCTION F_FloorDN : DINT
(*
Rounding down function which returns the biggest double integer.

Constructor: 		Patryk Panylo
Company:		E. Riexinger GmbH
Date:			20.01.2014
Version:			1.00

Date:			Revision:		Who:				Comment
dd.mm.yyyy		x.xx			Initials			comment

*)
VAR_INPUT
	rInValue						:REAL;
END_VAR
VAR
END_VAR


F_FloorDN := REAL_TO_DINT(rInValue);

IF DINT_TO_REAL(F_FloorDN) > rInValue
THEN
	F_FloorDN := F_FloorDN - 1;
END_IF

END_FUNCTION

// ---- POUs/Tc2 Objects/Mathematical/F_FracR.TcPOU
FUNCTION F_FracR : REAL
(*
Function used to get fraction part of a real number.

Constructor: 		Patryk Panylo
Company:		E. Riexinger GmbH
Date:			17.07.2014
Version:			1.00

Date:			Revision:		Who:				Comment
dd.mm.yyyy		x.xx			Initials			comment

*)
VAR_INPUT
	(* Enummerations *)

	(* Variables *)
	rReal 						:REAL;			(* Input variable *)

	(* References *)

	(* Interfaces *)

	(* Instances *)

END_VAR
VAR
	(* Enummerations *)
	
	(* Variables *)
	rFloor						:REAL;

	(* References *)

	(* Interfaces *)

	(* Instances *)

END_VAR


rFloor := DINT_TO_REAL(F_FloorDN(ABS(rReal)));								(* Floor the value *)

IF rReal < 0
THEN
	F_FracR := rReal + rFloor ;								(* The fraction of the value *)

ELSE
	F_FracR := rReal - rFloor;								(* The fraction of the value *)

END_IF

END_FUNCTION

// ---- POUs/Tc2 Objects/Mathematical/F_GCD.TcPOU
FUNCTION F_GCD : INT
(* Greatest common divisor *)
VAR_INPUT
	A : DINT;
	B : DINT;
END_VAR
VAR
	t: DINT;
END_VAR


(*
version 1.0	19. jan. 2011
programmer 	hugo
tested by	tobias

this function calculates the gretaest common divisor of two numbers A and B

*)

IF A = 0 THEN
	F_GCD := DINT_TO_INT(ABS(B));
ELSIF B = 0 THEN
	F_GCD := DINT_TO_INT(ABS(A));
ELSE
	A := ABS(A);
	B := ABS(B);
	F_GCD := 1;
	WHILE NOT(A.0 OR B.0) DO
		A := SHR(A,1);
		B := SHR(B,1);
		F_GCD := SHL(F_GCD,1);
	END_WHILE;
	WHILE A > 0 DO
		IF NOT(A.0) THEN A := SHR(A,1);
		ELSIF NOT(B.0) THEN B := SHR(B,1);
		ELSE
			t:= SHR(ABS(A-B),1);
			IF A < B THEN B := t; ELSE A := T; END_IF;
		END_IF;
	END_WHILE;
	F_GCD := F_GCD * DINT_TO_INT(B);
END_IF;


(* revision history
hm	19. jan. 2011	rev 1.0
	original version

*)

END_FUNCTION

// ---- POUs/Tc2 Objects/Mathematical/F_MM_TO_DEG.TcPOU
FUNCTION F_MM_TO_DEG : LREAL
(*

The function used to convert mm to deg.

Constructor: 		Patryk Panylo
Company:		E. Riexinger GmbH
Date:			12.11.2019
Version:			1.00

Date:			Revision:		Who:				Comment
dd.mm.yyyy		x.xx			Initials			comment

*)
VAR_INPUT
	(* Input variables / Eingang Variablen *)
	lrDiameter							:LREAL; 						(*  Input variable *)
	lrDistance							:LREAL; 						(*  Input variable *)
END_VAR
VAR
	(* Variables *)

END_VAR
VAR CONSTANT
	lrRotation							:LREAL := 360.0;				(* Rotation deg *)
END_VAR


IF lrDiameter <> 0
THEN
	F_MM_TO_DEG := lrDistance * lrRotation / (lrDiameter * PI);
ELSE
	F_MM_TO_DEG := 0.0;
END_IF

END_FUNCTION

// ---- POUs/Tc2 Objects/Mathematical/F_ModR.TcPOU
FUNCTION F_ModR : REAL
(*
Modulo function for real numbers (dividend mod divisor).

Constructor: 		Patryk Panylo
Company:		E. Riexinger GmbH
Date:			20.01.2014
Version:			1.00

Date:			Revision:		Who:				Comment
dd.mm.yyyy		x.xx			Initials			comment

*)
VAR_INPUT
	rDividend						:REAL;
	rDivisor							:REAL := 1.0;
END_VAR
VAR
END_VAR


F_ModR := rDivisor;

IF rDivisor <> 0.0 
THEN
	F_ModR := rDividend - DINT_TO_REAL(F_FloorDN(rDividend / rDivisor)) * rDivisor;
END_IF;

END_FUNCTION

// ---- POUs/Tc2 Objects/Mathematical/F_RoundR.TcPOU
FUNCTION F_RoundR : REAL
(*
Function used to round real value with precision

Constructor: 		Patryk Panylo
Company:		E. Riexinger GmbH
Date:			17.07.2014
Version:			1.00

Date:			Revision:		Who:				Comment
dd.mm.yyyy		x.xx			Initials			comment

*)
VAR_INPUT
	(* Enummerations *)
	
	(* Variables *)
	rReal 						:REAL;			(* Input variable *)
	usnPrecision					:USINT := 2;		(* The number of digits after the decimal point depends on the requested precision *)

	(* References *)

	(* Interfaces *)

	(* Instances *)

END_VAR
VAR
	(* Enummerations *)
	
	(* Variables *)
	rFraction						:REAL;

	(* References *)

	(* Interfaces *)

	(* Instances *)

END_VAR


rFraction := F_FracR(ABS(rReal)) * EXPT(10, usnPrecision + 1); 								(* The fraction of the value *)

IF F_ModR(rFraction, 10) < 5
THEN
	rFraction := rFraction - F_ModR(rFraction, 10) ;											(* Round down *)
ELSE
	rFraction := rFraction + (10 - F_ModR(rFraction, 10));										(* Round up and check the integral increment *)
END_IF;

IF rReal  < 0																			(* Check the digit of the value *)
THEN
	F_RoundR := TRUNC(rReal) - (rFraction / EXPT(10, usnPrecision + 1));
ELSE
	F_RoundR := TRUNC(rReal) + (rFraction / EXPT(10, usnPrecision + 1));
END_IF

END_FUNCTION

// ---- POUs/Tc2 Objects/Mathematical/Hysteresis/FB_Hysteresis.TcPOU
FUNCTION_BLOCK FB_Hysteresis
(*
Function block used to generate hysteresis

Constructor: 		Patryk Panylo
Company:		E. Riexinger GmbH
Date:			15.07.2016
Version:			1.00

Date:			Revision:		Who:				Comment
dd.mm.yyyy		x.xx			Initials			comment

*)
VAR_INPUT
	(* Enummerations *)

	(* Variables *)
	bEnable							:BOOL := TRUE;					(* Enable FB *)

	lrInSignal							:LREAL;							(* Input signal *)
	lrGoDown						:REAL;
	lrGoUp							:REAL;

	(* References *)

	(* Interfaces *)

	(* Instances *)
END_VAR
VAR_OUTPUT
	(* Enummerations *)
	
	(* Variables *)
	lrOutSignal						:LREAL;						(* Output signal *)
	bLowLevel						:BOOL;						(* Low level detected *)
	bGoLevel						:BOOL;						(* Go level detected *)
	bHighLevel						:BOOL;						(* High level detected *)

	(* References *)

	(* Interfaces *)

	(* Instances *)
END_VAR
VAR
	(* Enummerations *)

	(* Variables *)
	bFirstTime							:BOOL;							(* First cycle *)

	lrLastSignal							:LREAL;							(* Last signal *)

	(* References *)

	(* Interfaces *)

	(* Instances *)

END_VAR

IF NOT bEnable
THEN
	lrOutSignal := lrInSignal;

	bFirstTime := FALSE;
	RETURN;
END_IF

IF NOT bFirstTime
THEN

	bFirstTime := TRUE;
END_IF

lrOutSignal:=SEL(lrInSignal - lrGoUp > lrLastSignal, lrOutSignal, lrInSignal - lrGoUp);
lrOutSignal:=SEL(lrInSignal + lrGoDown < lrLastSignal, lrOutSignal, lrInSignal + lrGoDown);

lrLastSignal := lrOutSignal;

END_FUNCTION_BLOCK

// ---- POUs/Tc2 Objects/Mathematical/Limits/FB_Limiter.TcPOU
FUNCTION_BLOCK FB_Limiter
(*
Function block used to limits input signal. 

Constructor: 		Patryk Panylo
Company:		E. Riexinger GmbH
Date:			21.07.2014
Version:			1.00

Date:			Revision:		Who:				Comment
dd.mm.yyyy		x.xx			Initials			comment

*)
VAR_INPUT
	(* Enummerations *)

	(* Variables *)
	bEnable								:BOOL := TRUE;					(* Enable FB *)

	lrInSignal								:LREAL;							(* Input signal *)
	lrLimitMin								:LREAL;							(* Limit minimum *)
	lrLimitMax							:LREAL;							(* Limit maximum *)

	(* References *)

	(* Interfaces *)

	(* Instances *)
END_VAR
VAR_OUTPUT
	(* Enummerations *)
	
	(* Variables *)
	lrOutSignal							:LREAL;							(* Output signal *)
	bLimitMin							:BOOL;							(* Minimum limit reached *)
	bLimitMax							:BOOL;							(* Maximum limit reached *)

	(* References *)

	(* Interfaces *)

	(* Instances *)
END_VAR
VAR
	(* Enummerations *)
	
	(* Variables *)
	bFirstTime							:BOOL;							(* First cycle *)

	(* References *)

	(* Interfaces *)

	(* Instances *)

END_VAR

IF NOT bEnable
THEN
	lrOutSignal := lrInSignal;

	bLimitMin := FALSE;							(* Minimum limit reached *)
	bLimitMax := FALSE;							(* Maximum limit reached *)

	bFirstTime := FALSE;
	RETURN;
END_IF

IF NOT bFirstTime
THEN

	bFirstTime := TRUE;
END_IF

lrOutSignal := lrInSignal;
bLimitMin := FALSE;							(* Minimum limit reached *)
bLimitMax := FALSE;							(* Maximum limit reached *)

IF lrInSignal <= lrLimitMin
THEN
	lrOutSignal  := lrLimitMin;
	bLimitMin := TRUE;

ELSIF lrInSignal >= lrLimitMax
THEN
	lrOutSignal := lrLimitMax;
	bLimitMax := TRUE;

END_IF

END_FUNCTION_BLOCK

// ---- POUs/Tc2 Objects/Mathematical/Limits/F_DeadZone.TcPOU
FUNCTION F_DeadZone : REAL
(*
Function used to calculate dead zone.

Constructor: 		Patryk Panylo
Company:		E. Riexinger GmbH
Date:			03.06.2014
Version:			1.00

Date:			Revision:		Who:				Comment
dd.mm.yyyy		x.xx			Initials			comment

*)

VAR_INPUT
	(* Enummerations *)

	(* Variables *)
	lrInSignal								:LREAL;							(* Input signal *)
	lrDeadZone							:LREAL;							(* Dead zone *)

	(* References *)

	(* Interfaces *)

	(* Instances *)

END_VAR
VAR
	(* Enummerations *)

	(* Variables *)

	(* References *)

	(* Interfaces *)

	(* Instances *)

END_VAR


IF ABS(lrInSignal) > lrDeadZone
THEN
	F_DeadZone := lrInSignal;
ELSE
	F_DeadZone := 0.0;
END_IF;

END_FUNCTION

// ---- POUs/Tc2 Objects/Mathematical/Limits/F_WordToRange.TcPOU
FUNCTION F_WordToRange : REAL
VAR_INPUT
	wWord 					:WORD;
	rLowLimit 				:REAL;
	rHighLimit 				:REAL;
END_VAR
VAR
END_VAR


F_WordToRange := (rHighLimit - rLowLimit) * WORD_TO_REAL(wWord) * 0.00001525902189669640 + rLowLimit;

END_FUNCTION

// ---- POUs/Tc2 Objects/Measurements/Counter/FB_DistanceCounter.TcPOU
FUNCTION_BLOCK FB_DistanceCounter
(*

Function block to read and write elapsed distance in/from file.
If sFileName or sFilePath  or sFileSuffix is empty then save function is diabled and generate error.

Constructor: 		Patryk Panylo
Company:		E. Riexinger GmbH
Date:			24.03.2014
Version:			1.00

Date:			Revision:		Who:				Comment
dd.mm.yyyy		x.xx			Initials			comment

*)

VAR_INPUT
	(* Variables *)
	bEnable							:BOOL;							(* Enable FB *)
	sAmsNetId 						:STRING := ''; 						(* Ams Net ID of file to read/write *)
	lrDistance						:LREAL; 							(* All over counter distance *)
	bCount							:BOOL; 							(* If true then count distance else save current distance *)
	bSave							:BOOL;							(* Save current distance counter *)
	bReset							:BOOL; 							(* Reset counter *)
	bDeleteAll						:BOOL; 							(* Delete all counters since beginning *)
	sFilePath						:STRING := 'C:\TwinCAT\Plc\';		(* File path *)
	sFileName						:STRING := 'default';				(* File name *)
	tSaveIntervall						:TIME := t#3m;						(* Intervall to save counter hours. If equal 0 then intervall is off *)
	tTimeout							:TIME := t#3s;						(* ADS timeout *)
END_VAR
VAR_OUTPUT
	(* Variables *)
	lrAllOverDistance					:LREAL; 							(* All over counter distance *)
	lrAfterResetDistance				:LREAL; 							(* Counter distance since last reset *)
	lrNoRetainDistance				:LREAL; 							(* No retain counter distance *)
	bError							:BOOL;							(* Program error *)
	udnErrNo						:UDINT;							(* Error number *)
END_VAR
VAR
	(* Enummerations *)
	etRWStep						:(eReadDistance, eChkRead, eWFWrite, eWriteDistance, eChkWrite, eError );

	(* Variables *)
	bFirstTime						:BOOL;
	stRetainDistance					:ST_DistanceCounter;
	stCacheRetainDistance			:ST_DistanceCounter;

	(* Instances *)
	ftCount							:F_TRIG;
	rtSave							:R_TRIG;
	rtReset							:R_TRIG;
	rtDeleteAll						:R_TRIG;

	fbFileHandler						:FB_FileHandlerBinary;				(* File handler *)
	tonWriteIntervall					:TON;							(* Timer for Save intervall control *)

END_VAR

IF NOT bEnable				(* Enable FB *)
THEN
	fbFileHandler(
		bEnable := FALSE,
		bExecute := FALSE,
		bFileRead := FALSE,
		bFileWrite := FALSE
	);

	bFirstTime := FALSE;
	bError := FALSE;			(* Program error *)
	udnErrNo := 0;				(* Error number *)

	RETURN;
END_IF


IF NOT bFirstTime
THEN
	(* Produce the file directory name *)
	fbFileHandler.sFilePath := sFilePath;
	fbFileHandler.sFileName := sFileName;
	fbFileHandler.sFileSuffix := 'dc';

	tonWriteIntervall(
		IN := FALSE,
		PT:= tSaveIntervall
	);

	etRWStep := eReadDistance;

	bFirstTime := TRUE;
	RETURN;
END_IF


(* Read / Write all over distance *)
CASE etRWStep OF

	eReadDistance:
		fbFileHandler.bExecute := TRUE;
		fbFileHandler.bFileRead := TRUE;
		fbFileHandler.bFileWrite := FALSE;

		IF fbFileHandler.bBusy
		THEN
			etRWStep := eChkRead;

		END_IF

	eChkRead:
		IF NOT fbFileHandler.bBusy
		THEN
			IF  fbFileHandler.bError
			THEN
				fbFileHandler.bExecute := FALSE;
				fbFileHandler.bFileRead := FALSE;
				fbFileHandler.bFileWrite := FALSE;

				stCacheRetainDistance.lrAllOverDistance := 0;
				stCacheRetainDistance.lrAfterResetDistance := 0;

				etRWStep := eWFWrite;				(* Next step *)

			ELSE
				fbFileHandler.bExecute := FALSE;
				fbFileHandler.bFileRead := FALSE;
				fbFileHandler.bFileWrite := FALSE;

				stCacheRetainDistance.lrAllOverDistance := stRetainDistance.lrAllOverDistance;
				stCacheRetainDistance.lrAfterResetDistance := stRetainDistance.lrAfterResetDistance;

				etRWStep := eWFWrite;				(* Next step *)

			END_IF
		END_IF

	eWFWrite:
		ftCount(
			CLK :=  bCount AND NOT bReset AND NOT bDeleteAll
		);

		rtSave(
			CLK := bSave AND NOT bReset AND NOT bDeleteAll
		);


		tonWriteIntervall(IN := tSaveIntervall > t#0s);

		IF ftCount.Q
		     OR rtSave.Q
		     OR tonWriteIntervall.Q
		THEN
			tonWriteIntervall(IN := FALSE);

			etRWStep := eWriteDistance;								(* Next step *)

		END_IF

	eWriteDistance:
		fbFileHandler.bExecute := TRUE;
		fbFileHandler.bFileRead := FALSE;
		fbFileHandler.bFileWrite := TRUE;

		IF fbFileHandler.bBusy
		THEN
			etRWStep := eChkWrite;								(* Next step *)

		END_IF

	eChkWrite:
		IF NOT fbFileHandler.bBusy
		THEN
			IF  fbFileHandler.bError
			THEN
				etRWStep := eError;								(* Next step *)

			ELSE
				fbFileHandler.bExecute := FALSE;
				fbFileHandler.bFileRead := FALSE;
				fbFileHandler.bFileWrite := FALSE;

				etRWStep := eWFWrite;							(* Next step *)

			END_IF
		END_IF

	eError:
		fbFileHandler.bExecute := FALSE;
		fbFileHandler.bFileRead := FALSE;
		fbFileHandler.bFileWrite := FALSE;

END_CASE


